{region "02 - Accept Start"}
// Accept Start into Starting; processing and Assertion evaluation are not active yet.
FSteps[2].RequestStart := TRUE;
FSteps[2].ExpectedState := E_State.Starting;
FSteps[2].ExpectedResult := E_Result.NotEvaluated;
FSteps[2].ExpectedReady := FALSE;
FSteps[2].ExpectedPassedCount := 0;
FSteps[2].ExpectedFailedCount := 0;
FSteps[2].ExpectedHookCount := 5;
FSteps[2].ExpectedHooks[1].Hook := E_LifecycleHook.Abort;
FSteps[2].ExpectedHooks[1].State := E_State.Starting;
FSteps[2].ExpectedHooks[1].Enabled := FALSE;
FSteps[2].ExpectedHooks[2].Hook := E_LifecycleHook.Preparations;
FSteps[2].ExpectedHooks[2].State := E_State.Starting;
FSteps[2].ExpectedHooks[2].Enabled := FALSE;
FSteps[2].ExpectedHooks[3].Hook := E_LifecycleHook.Tests;
FSteps[2].ExpectedHooks[3].State := E_State.Starting;
FSteps[2].ExpectedHooks[3].Enabled := FALSE;
FSteps[2].ExpectedHooks[4].Hook := E_LifecycleHook.Assertions;
FSteps[2].ExpectedHooks[4].State := E_State.Starting;
FSteps[2].ExpectedHooks[4].Enabled := FALSE;
FSteps[2].ExpectedHooks[5].Hook := E_LifecycleHook.Aggregate;
FSteps[2].ExpectedHooks[5].State := E_State.Starting;
FSteps[2].ExpectedHooks[5].Enabled := TRUE;
{endregion}

{region "03 - Enter Running"}
// Enter Running and evaluate both children; owner Result stays NotEvaluated until finalization.
FSteps[3].ExpectedState := E_State.Running;
FSteps[3].ExpectedResult := E_Result.NotEvaluated;
FSteps[3].ExpectedReady := FALSE;
FSteps[3].ExpectedPassedCount := 2;
FSteps[3].ExpectedFailedCount := 0;
FSteps[3].ExpectedHookCount := 5;
FSteps[3].ExpectedHooks[1].Hook := E_LifecycleHook.Abort;
FSteps[3].ExpectedHooks[1].State := E_State.Running;
FSteps[3].ExpectedHooks[1].Enabled := FALSE;
FSteps[3].ExpectedHooks[2].Hook := E_LifecycleHook.Preparations;
FSteps[3].ExpectedHooks[2].State := E_State.Running;
FSteps[3].ExpectedHooks[2].Enabled := FALSE;
FSteps[3].ExpectedHooks[3].Hook := E_LifecycleHook.Tests;
FSteps[3].ExpectedHooks[3].State := E_State.Running;
FSteps[3].ExpectedHooks[3].Enabled := TRUE;
FSteps[3].ExpectedHooks[4].Hook := E_LifecycleHook.Assertions;
FSteps[3].ExpectedHooks[4].State := E_State.Running;
FSteps[3].ExpectedHooks[4].Enabled := TRUE;
FSteps[3].ExpectedHooks[5].Hook := E_LifecycleHook.Aggregate;
FSteps[3].ExpectedHooks[5].State := E_State.Running;
FSteps[3].ExpectedHooks[5].Enabled := TRUE;
{endregion}

{region "04 - Request Abort and hold acknowledgement"}
// Request Abort once and withhold cleanup acknowledgement.
FSteps[4].RequestAbort := TRUE;
FSteps[4].AbortCompleted := FALSE;
FSteps[4].ExpectedState := E_State.Aborting;
FSteps[4].ExpectedResult := E_Result.Abort;
FSteps[4].ExpectedReady := FALSE;
FSteps[4].ExpectedPassedCount := 2;
FSteps[4].ExpectedFailedCount := 0;
FSteps[4].ExpectedHookCount := 5;
FSteps[4].ExpectedHooks[1].Hook := E_LifecycleHook.Abort;
FSteps[4].ExpectedHooks[1].State := E_State.Aborting;
FSteps[4].ExpectedHooks[1].Enabled := TRUE;
FSteps[4].ExpectedHooks[2].Hook := E_LifecycleHook.Preparations;
FSteps[4].ExpectedHooks[2].State := E_State.Aborting;
FSteps[4].ExpectedHooks[2].Enabled := FALSE;
FSteps[4].ExpectedHooks[3].Hook := E_LifecycleHook.Tests;
FSteps[4].ExpectedHooks[3].State := E_State.Aborting;
FSteps[4].ExpectedHooks[3].Enabled := FALSE;
FSteps[4].ExpectedHooks[4].Hook := E_LifecycleHook.Assertions;
FSteps[4].ExpectedHooks[4].State := E_State.Aborting;
FSteps[4].ExpectedHooks[4].Enabled := FALSE;
FSteps[4].ExpectedHooks[5].Hook := E_LifecycleHook.Aggregate;
FSteps[4].ExpectedHooks[5].State := E_State.Aborting;
FSteps[4].ExpectedHooks[5].Enabled := TRUE;
{endregion}

{region "05 - Wait for Abort timeout"}
// Keep cleanup open while repeating this checkpoint in Aborting.
// Timeout forces Completing with Error even though the implementation never acknowledges Abort.
FSteps[5].WaitForTransition := TRUE;
FSteps[5].WaitingState := E_State.Aborting;
FSteps[5].AbortCompleted := FALSE;
FSteps[5].ExpectedAbortTimeout := TRUE;
FSteps[5].ExpectedState := E_State.Completing;
FSteps[5].ExpectedResult := E_Result.Error;
FSteps[5].ExpectedReady := FALSE;
FSteps[5].ExpectedPassedCount := 2;
FSteps[5].ExpectedFailedCount := 0;
FSteps[5].ExpectedHookCount := 5;
FSteps[5].ExpectedHooks[1].Hook := E_LifecycleHook.Abort;
FSteps[5].ExpectedHooks[1].State := E_State.Completing;
FSteps[5].ExpectedHooks[1].Enabled := FALSE;
FSteps[5].ExpectedHooks[2].Hook := E_LifecycleHook.Preparations;
FSteps[5].ExpectedHooks[2].State := E_State.Completing;
FSteps[5].ExpectedHooks[2].Enabled := FALSE;
FSteps[5].ExpectedHooks[3].Hook := E_LifecycleHook.Tests;
FSteps[5].ExpectedHooks[3].State := E_State.Completing;
FSteps[5].ExpectedHooks[3].Enabled := FALSE;
FSteps[5].ExpectedHooks[4].Hook := E_LifecycleHook.Assertions;
FSteps[5].ExpectedHooks[4].State := E_State.Completing;
FSteps[5].ExpectedHooks[4].Enabled := FALSE;
FSteps[5].ExpectedHooks[5].Hook := E_LifecycleHook.Aggregate;
FSteps[5].ExpectedHooks[5].State := E_State.Completing;
FSteps[5].ExpectedHooks[5].Enabled := TRUE;
{endregion}

{region "06 - Retain timeout at completion"}
// Reach Completed and retain the Abort-timeout diagnostic.
FSteps[6].ExpectedAbortTimeout := TRUE;
FSteps[6].ExpectedState := E_State.Completed;
FSteps[6].ExpectedResult := E_Result.Error;
FSteps[6].ExpectedReady := FALSE;
FSteps[6].ExpectedPassedCount := 2;
FSteps[6].ExpectedFailedCount := 0;
FSteps[6].ExpectedHookCount := 1;
FSteps[6].ExpectedHooks[1].Hook := E_LifecycleHook.Aggregate;
FSteps[6].ExpectedHooks[1].State := E_State.Completed;
FSteps[6].ExpectedHooks[1].Enabled := TRUE;
{endregion}

{region "07 - Reset clears held timeout and result"}
FSteps[7].ExpectedState := E_State.Idle;
FSteps[7].ExpectedResult := E_Result.NotEvaluated;
FSteps[7].ExpectedReady := TRUE;
FSteps[7].ExpectedPassedCount := 0;
FSteps[7].ExpectedFailedCount := 0;
FSteps[7].CheckFinalization := TRUE;
FSteps[7].ExpectedFinalizationCount := 1;
FSteps[7].ExpectedCompletionCount := 1;
FSteps[7].ExpectedFinalResult := E_Result.Error;
FSteps[7].RequestReset := TRUE;
FSteps[7].PreparationTargetReached := TRUE;
FSteps[7].ExpectRuntimeCleared := TRUE;
FSteps[7].ExpectedHookCount := 6;
FSteps[7].ExpectedHooks[1].Hook := E_LifecycleHook.Reset;
FSteps[7].ExpectedHooks[1].State := E_State.Reset;
FSteps[7].ExpectedHooks[1].Enabled := TRUE;
FSteps[7].ExpectedHooks[2].Hook := E_LifecycleHook.Abort;
FSteps[7].ExpectedHooks[2].State := E_State.Idle;
FSteps[7].ExpectedHooks[2].Enabled := FALSE;
FSteps[7].ExpectedHooks[3].Hook := E_LifecycleHook.Preparations;
FSteps[7].ExpectedHooks[3].State := E_State.Idle;
FSteps[7].ExpectedHooks[3].Enabled := FALSE;
FSteps[7].ExpectedHooks[4].Hook := E_LifecycleHook.Tests;
FSteps[7].ExpectedHooks[4].State := E_State.Idle;
FSteps[7].ExpectedHooks[4].Enabled := FALSE;
FSteps[7].ExpectedHooks[5].Hook := E_LifecycleHook.Assertions;
FSteps[7].ExpectedHooks[5].State := E_State.Idle;
FSteps[7].ExpectedHooks[5].Enabled := FALSE;
FSteps[7].ExpectedHooks[6].Hook := E_LifecycleHook.Aggregate;
FSteps[7].ExpectedHooks[6].State := E_State.Idle;
FSteps[7].ExpectedHooks[6].Enabled := TRUE;
{endregion}

{region "08 - Start after timeout recovery"}
FSteps[8].ExpectedState := E_State.Starting;
FSteps[8].ExpectedResult := E_Result.NotEvaluated;
FSteps[8].ExpectedReady := FALSE;
FSteps[8].ExpectedPassedCount := 0;
FSteps[8].ExpectedFailedCount := 0;
FSteps[8].CheckFinalization := TRUE;
FSteps[8].ExpectedFinalizationCount := 1;
FSteps[8].ExpectedCompletionCount := 1;
FSteps[8].ExpectedFinalResult := E_Result.Error;
FSteps[8].RequestStart := TRUE;
FSteps[8].PreparationTargetReached := TRUE;
FSteps[8].ExpectedHookCount := 5;
FSteps[8].ExpectedHooks[1].Hook := E_LifecycleHook.Abort;
FSteps[8].ExpectedHooks[1].State := E_State.Starting;
FSteps[8].ExpectedHooks[1].Enabled := FALSE;
FSteps[8].ExpectedHooks[2].Hook := E_LifecycleHook.Preparations;
FSteps[8].ExpectedHooks[2].State := E_State.Starting;
FSteps[8].ExpectedHooks[2].Enabled := FALSE;
FSteps[8].ExpectedHooks[3].Hook := E_LifecycleHook.Tests;
FSteps[8].ExpectedHooks[3].State := E_State.Starting;
FSteps[8].ExpectedHooks[3].Enabled := FALSE;
FSteps[8].ExpectedHooks[4].Hook := E_LifecycleHook.Assertions;
FSteps[8].ExpectedHooks[4].State := E_State.Starting;
FSteps[8].ExpectedHooks[4].Enabled := FALSE;
FSteps[8].ExpectedHooks[5].Hook := E_LifecycleHook.Aggregate;
FSteps[8].ExpectedHooks[5].State := E_State.Starting;
FSteps[8].ExpectedHooks[5].Enabled := TRUE;
{endregion}

{region "09 - Execute without previous timeout flags"}
FSteps[9].ExpectedState := E_State.Running;
FSteps[9].ExpectedResult := E_Result.NotEvaluated;
FSteps[9].ExpectedReady := FALSE;
FSteps[9].ExpectedPassedCount := 2;
FSteps[9].ExpectedFailedCount := 0;
FSteps[9].CheckFinalization := TRUE;
FSteps[9].ExpectedFinalizationCount := 1;
FSteps[9].ExpectedCompletionCount := 1;
FSteps[9].ExpectedFinalResult := E_Result.Error;
FSteps[9].ExpectedHookCount := 5;
FSteps[9].ExpectedHooks[1].Hook := E_LifecycleHook.Abort;
FSteps[9].ExpectedHooks[1].State := E_State.Running;
FSteps[9].ExpectedHooks[1].Enabled := FALSE;
FSteps[9].ExpectedHooks[2].Hook := E_LifecycleHook.Preparations;
FSteps[9].ExpectedHooks[2].State := E_State.Running;
FSteps[9].ExpectedHooks[2].Enabled := FALSE;
FSteps[9].ExpectedHooks[3].Hook := E_LifecycleHook.Tests;
FSteps[9].ExpectedHooks[3].State := E_State.Running;
FSteps[9].ExpectedHooks[3].Enabled := TRUE;
FSteps[9].ExpectedHooks[4].Hook := E_LifecycleHook.Assertions;
FSteps[9].ExpectedHooks[4].State := E_State.Running;
FSteps[9].ExpectedHooks[4].Enabled := TRUE;
FSteps[9].ExpectedHooks[5].Hook := E_LifecycleHook.Aggregate;
FSteps[9].ExpectedHooks[5].State := E_State.Running;
FSteps[9].ExpectedHooks[5].Enabled := TRUE;
{endregion}

{region "10 - Finalize the recovered run"}
FSteps[10].ExpectedState := E_State.Completing;
FSteps[10].ExpectedResult := E_Result.Passed;
FSteps[10].ExpectedReady := FALSE;
FSteps[10].ExpectedPassedCount := 2;
FSteps[10].ExpectedFailedCount := 0;
FSteps[10].FinishTests := TRUE;
FSteps[10].CheckFinalization := TRUE;
FSteps[10].ExpectedFinalizationCount := 2;
FSteps[10].ExpectedCompletionCount := 1;
FSteps[10].ExpectedFinalResult := E_Result.Passed;
FSteps[10].ExpectedHookCount := 5;
FSteps[10].ExpectedHooks[1].Hook := E_LifecycleHook.Abort;
FSteps[10].ExpectedHooks[1].State := E_State.Running;
FSteps[10].ExpectedHooks[1].Enabled := FALSE;
FSteps[10].ExpectedHooks[2].Hook := E_LifecycleHook.Preparations;
FSteps[10].ExpectedHooks[2].State := E_State.Running;
FSteps[10].ExpectedHooks[2].Enabled := FALSE;
FSteps[10].ExpectedHooks[3].Hook := E_LifecycleHook.Tests;
FSteps[10].ExpectedHooks[3].State := E_State.Running;
FSteps[10].ExpectedHooks[3].Enabled := TRUE;
FSteps[10].ExpectedHooks[4].Hook := E_LifecycleHook.Assertions;
FSteps[10].ExpectedHooks[4].State := E_State.Completing;
FSteps[10].ExpectedHooks[4].Enabled := FALSE;
FSteps[10].ExpectedHooks[5].Hook := E_LifecycleHook.Aggregate;
FSteps[10].ExpectedHooks[5].State := E_State.Completing;
FSteps[10].ExpectedHooks[5].Enabled := TRUE;
{endregion}

{region "11 - Complete the recovered run"}
FSteps[11].ExpectedState := E_State.Completed;
FSteps[11].ExpectedResult := E_Result.Passed;
FSteps[11].ExpectedReady := FALSE;
FSteps[11].ExpectedPassedCount := 2;
FSteps[11].ExpectedFailedCount := 0;
FSteps[11].ExpectRuntimeHeld := TRUE;
FSteps[11].CheckFinalization := TRUE;
FSteps[11].ExpectedFinalizationCount := 2;
FSteps[11].ExpectedCompletionCount := 2;
FSteps[11].ExpectedFinalResult := E_Result.Passed;
FSteps[11].ExpectedHookCount := 1;
FSteps[11].ExpectedHooks[1].Hook := E_LifecycleHook.Aggregate;
FSteps[11].ExpectedHooks[1].State := E_State.Completed;
FSteps[11].ExpectedHooks[1].Enabled := TRUE;
{endregion}

{region "12 - Hold the recovered completion without new events"}
FSteps[12].ExpectedState := E_State.Completed;
FSteps[12].ExpectedResult := E_Result.Passed;
FSteps[12].ExpectedReady := FALSE;
FSteps[12].ExpectedPassedCount := 2;
FSteps[12].ExpectedFailedCount := 0;
FSteps[12].ExpectQuietCall := TRUE;
FSteps[12].ExpectRuntimeHeld := TRUE;
FSteps[12].CheckFinalization := TRUE;
FSteps[12].ExpectedFinalizationCount := 2;
FSteps[12].ExpectedCompletionCount := 2;
FSteps[12].ExpectedFinalResult := E_Result.Passed;
FSteps[12].ExpectedHookCount := 1;
FSteps[12].ExpectedHooks[1].Hook := E_LifecycleHook.Aggregate;
FSteps[12].ExpectedHooks[1].State := E_State.Completed;
FSteps[12].ExpectedHooks[1].Enabled := TRUE;
{endregion}
END_METHOD

END_FUNCTION_BLOCK

// ---- SelfTests/TestCases/TestSuite_TestCaseLifecycle/Test_LifecycleExecutionTimeout.TcPOU
{region 'Documentation'}
(*!
<summary>Leaves the Test phase pending until the real configured execution timeout finalizes Error.</summary>
*)
{endregion}
FUNCTION_BLOCK Test_LifecycleExecutionTimeout EXTENDS TestCaseLifecycleTestBase

SUPER^();

{region 'Documentation'}
(*!
<summary>Defines explicit exceptional-path stimuli and contract-derived observations.</summary>
*)
{endregion}
METHOD PROTECTED ConfigureScenario
// Exercise the real cyclic timer; these checkpoints check the timeout path and retained flag,
// not an exact elapsed-time boundary. The outer Test Case timeout bounds a missing transition.
FSubjectPreparationCount := 0;
FSubjectTestCount := 1;
FStepCount := 11;
FSubjectConfig.Timeout := T#50ms;

{region "01 - Reset to Idle"}
// Establish Idle through the parent Reset request; both child results must be cleared.
FSteps[1].RequestReset := TRUE;
FSteps[1].ExpectedState := E_State.Idle;
FSteps[1].ExpectedResult := E_Result.NotEvaluated;
FSteps[1].ExpectedReady := TRUE;
FSteps[1].ExpectedPassedCount := 0;
FSteps[1].ExpectedFailedCount := 0;
FSteps[1].ExpectedHookCount := 6;
FSteps[1].ExpectedHooks[1].Hook := E_LifecycleHook.Reset;
FSteps[1].ExpectedHooks[1].State := E_State.Reset;
FSteps[1].ExpectedHooks[1].Enabled := TRUE;
FSteps[1].ExpectedHooks[2].Hook := E_LifecycleHook.Abort;
FSteps[1].ExpectedHooks[2].State := E_State.Idle;
FSteps[1].ExpectedHooks[2].Enabled := FALSE;
FSteps[1].ExpectedHooks[3].Hook := E_LifecycleHook.Preparations;
FSteps[1].ExpectedHooks[3].State := E_State.Idle;
FSteps[1].ExpectedHooks[3].Enabled := FALSE;
FSteps[1].ExpectedHooks[4].Hook := E_LifecycleHook.Tests;
FSteps[1].ExpectedHooks[4].State := E_State.Idle;
FSteps[1].ExpectedHooks[4].Enabled := FALSE;
FSteps[1].ExpectedHooks[5].Hook := E_LifecycleHook.Assertions;
FSteps[1].ExpectedHooks[5].State := E_State.Idle;
FSteps[1].ExpectedHooks[5].Enabled := FALSE;
FSteps[1].ExpectedHooks[6].Hook := E_LifecycleHook.Aggregate;
FSteps[1].ExpectedHooks[6].State := E_State.Idle;
FSteps[1].ExpectedHooks[6].Enabled := TRUE;
{endregion}

{region "02 - Accept Start"}
// Accept Start into Starting; processing and Assertion evaluation are not active yet.
FSteps[2].RequestStart := TRUE;
FSteps[2].ExpectedState := E_State.Starting;
FSteps[2].ExpectedResult := E_Result.NotEvaluated;
FSteps[2].ExpectedReady := FALSE;
FSteps[2].ExpectedPassedCount := 0;
FSteps[2].ExpectedFailedCount := 0;
FSteps[2].ExpectedHookCount := 5;
FSteps[2].ExpectedHooks[1].Hook := E_LifecycleHook.Abort;
FSteps[2].ExpectedHooks[1].State := E_State.Starting;
FSteps[2].ExpectedHooks[1].Enabled := FALSE;
FSteps[2].ExpectedHooks[2].Hook := E_LifecycleHook.Preparations;
FSteps[2].ExpectedHooks[2].State := E_State.Starting;
FSteps[2].ExpectedHooks[2].Enabled := FALSE;
FSteps[2].ExpectedHooks[3].Hook := E_LifecycleHook.Tests;
FSteps[2].ExpectedHooks[3].State := E_State.Starting;
FSteps[2].ExpectedHooks[3].Enabled := FALSE;
FSteps[2].ExpectedHooks[4].Hook := E_LifecycleHook.Assertions;
FSteps[2].ExpectedHooks[4].State := E_State.Starting;
FSteps[2].ExpectedHooks[4].Enabled := FALSE;
FSteps[2].ExpectedHooks[5].Hook := E_LifecycleHook.Aggregate;
FSteps[2].ExpectedHooks[5].State := E_State.Starting;
FSteps[2].ExpectedHooks[5].Enabled := TRUE;
{endregion}

{region "03 - Enter Running"}
// Enter Running and evaluate both children; owner Result stays NotEvaluated until finalization.
FSteps[3].ExpectedState := E_State.Running;
FSteps[3].ExpectedResult := E_Result.NotEvaluated;
FSteps[3].ExpectedReady := FALSE;
FSteps[3].ExpectedPassedCount := 2;
FSteps[3].ExpectedFailedCount := 0;
FSteps[3].ExpectedHookCount := 5;
FSteps[3].ExpectedHooks[1].Hook := E_LifecycleHook.Abort;
FSteps[3].ExpectedHooks[1].State := E_State.Running;
FSteps[3].ExpectedHooks[1].Enabled := FALSE;
FSteps[3].ExpectedHooks[2].Hook := E_LifecycleHook.Preparations;
FSteps[3].ExpectedHooks[2].State := E_State.Running;
FSteps[3].ExpectedHooks[2].Enabled := FALSE;
FSteps[3].ExpectedHooks[3].Hook := E_LifecycleHook.Tests;
FSteps[3].ExpectedHooks[3].State := E_State.Running;
FSteps[3].ExpectedHooks[3].Enabled := TRUE;
FSteps[3].ExpectedHooks[4].Hook := E_LifecycleHook.Assertions;
FSteps[3].ExpectedHooks[4].State := E_State.Running;
FSteps[3].ExpectedHooks[4].Enabled := TRUE;
FSteps[3].ExpectedHooks[5].Hook := E_LifecycleHook.Aggregate;
FSteps[3].ExpectedHooks[5].State := E_State.Running;
FSteps[3].ExpectedHooks[5].Enabled := TRUE;
{endregion}

{region "04 - Wait for execution timeout"}
// Keep execution open and repeat this checkpoint while Running.
// On timeout, immediate abort cleanup reaches Completing with Error and HasTimeout set.
FSteps[4].WaitForTransition := TRUE;
FSteps[4].WaitingState := E_State.Running;
FSteps[4].ExpectedTimeout := TRUE;
FSteps[4].ExpectedState := E_State.Completing;
FSteps[4].ExpectedResult := E_Result.Error;
FSteps[4].ExpectedReady := FALSE;
FSteps[4].ExpectedPassedCount := 2;
FSteps[4].ExpectedFailedCount := 0;
FSteps[4].ExpectedHookCount := 5;
FSteps[4].ExpectedHooks[1].Hook := E_LifecycleHook.Abort;
FSteps[4].ExpectedHooks[1].State := E_State.AbortingFromError;
FSteps[4].ExpectedHooks[1].Enabled := TRUE;
FSteps[4].ExpectedHooks[2].Hook := E_LifecycleHook.Preparations;
FSteps[4].ExpectedHooks[2].State := E_State.Completing;
FSteps[4].ExpectedHooks[2].Enabled := FALSE;
FSteps[4].ExpectedHooks[3].Hook := E_LifecycleHook.Tests;
FSteps[4].ExpectedHooks[3].State := E_State.Completing;
FSteps[4].ExpectedHooks[3].Enabled := FALSE;
FSteps[4].ExpectedHooks[4].Hook := E_LifecycleHook.Assertions;
FSteps[4].ExpectedHooks[4].State := E_State.Completing;
FSteps[4].ExpectedHooks[4].Enabled := FALSE;
FSteps[4].ExpectedHooks[5].Hook := E_LifecycleHook.Aggregate;
FSteps[4].ExpectedHooks[5].State := E_State.Completing;
FSteps[4].ExpectedHooks[5].Enabled := TRUE;
{endregion}

{region "05 - Retain timeout at completion"}
// Reach Completed and retain the execution-timeout diagnostic.
FSteps[5].ExpectedTimeout := TRUE;
FSteps[5].ExpectedState := E_State.Completed;
FSteps[5].ExpectedResult := E_Result.Error;
FSteps[5].ExpectedReady := FALSE;
FSteps[5].ExpectedPassedCount := 2;
FSteps[5].ExpectedFailedCount := 0;
FSteps[5].ExpectedHookCount := 1;
FSteps[5].ExpectedHooks[1].Hook := E_LifecycleHook.Aggregate;
FSteps[5].ExpectedHooks[1].State := E_State.Completed;
FSteps[5].ExpectedHooks[1].Enabled := TRUE;
{endregion}

{region "06 - Reset clears held timeout and result"}
FSteps[6].ExpectedState := E_State.Idle;
FSteps[6].ExpectedResult := E_Result.NotEvaluated;
FSteps[6].ExpectedReady := TRUE;
FSteps[6].ExpectedPassedCount := 0;
FSteps[6].ExpectedFailedCount := 0;
FSteps[6].CheckFinalization := TRUE;
FSteps[6].ExpectedFinalizationCount := 1;
FSteps[6].ExpectedCompletionCount := 1;
FSteps[6].ExpectedFinalResult := E_Result.Error;
FSteps[6].RequestReset := TRUE;
FSteps[6].PreparationTargetReached := TRUE;
FSteps[6].ExpectRuntimeCleared := TRUE;
FSteps[6].ExpectedHookCount := 6;
FSteps[6].ExpectedHooks[1].Hook := E_LifecycleHook.Reset;
FSteps[6].ExpectedHooks[1].State := E_State.Reset;
FSteps[6].ExpectedHooks[1].Enabled := TRUE;
FSteps[6].ExpectedHooks[2].Hook := E_LifecycleHook.Abort;
FSteps[6].ExpectedHooks[2].State := E_State.Idle;
FSteps[6].ExpectedHooks[2].Enabled := FALSE;
FSteps[6].ExpectedHooks[3].Hook := E_LifecycleHook.Preparations;
FSteps[6].ExpectedHooks[3].State := E_State.Idle;
FSteps[6].ExpectedHooks[3].Enabled := FALSE;
FSteps[6].ExpectedHooks[4].Hook := E_LifecycleHook.Tests;
FSteps[6].ExpectedHooks[4].State := E_State.Idle;
FSteps[6].ExpectedHooks[4].Enabled := FALSE;
FSteps[6].ExpectedHooks[5].Hook := E_LifecycleHook.Assertions;
FSteps[6].ExpectedHooks[5].State := E_State.Idle;
FSteps[6].ExpectedHooks[5].Enabled := FALSE;
FSteps[6].ExpectedHooks[6].Hook := E_LifecycleHook.Aggregate;
FSteps[6].ExpectedHooks[6].State := E_State.Idle;
FSteps[6].ExpectedHooks[6].Enabled := TRUE;
{endregion}

{region "07 - Start after timeout recovery"}
FSteps[7].ExpectedState := E_State.Starting;
FSteps[7].ExpectedResult := E_Result.NotEvaluated;
FSteps[7].ExpectedReady := FALSE;
FSteps[7].ExpectedPassedCount := 0;
FSteps[7].ExpectedFailedCount := 0;
FSteps[7].CheckFinalization := TRUE;
FSteps[7].ExpectedFinalizationCount := 1;
FSteps[7].ExpectedCompletionCount := 1;
FSteps[7].ExpectedFinalResult := E_Result.Error;
FSteps[7].RequestStart := TRUE;
FSteps[7].PreparationTargetReached := TRUE;
FSteps[7].ExpectedHookCount := 5;
FSteps[7].ExpectedHooks[1].Hook := E_LifecycleHook.Abort;
FSteps[7].ExpectedHooks[1].State := E_State.Starting;
FSteps[7].ExpectedHooks[1].Enabled := FALSE;
FSteps[7].ExpectedHooks[2].Hook := E_LifecycleHook.Preparations;
FSteps[7].ExpectedHooks[2].State := E_State.Starting;
FSteps[7].ExpectedHooks[2].Enabled := FALSE;
FSteps[7].ExpectedHooks[3].Hook := E_LifecycleHook.Tests;
FSteps[7].ExpectedHooks[3].State := E_State.Starting;
FSteps[7].ExpectedHooks[3].Enabled := FALSE;
FSteps[7].ExpectedHooks[4].Hook := E_LifecycleHook.Assertions;
FSteps[7].ExpectedHooks[4].State := E_State.Starting;
FSteps[7].ExpectedHooks[4].Enabled := FALSE;
FSteps[7].ExpectedHooks[5].Hook := E_LifecycleHook.Aggregate;
FSteps[7].ExpectedHooks[5].State := E_State.Starting;
FSteps[7].ExpectedHooks[5].Enabled := TRUE;
{endregion}

{region "08 - Execute without previous timeout flags"}
FSteps[8].ExpectedState := E_State.Running;
FSteps[8].ExpectedResult := E_Result.NotEvaluated;
FSteps[8].ExpectedReady := FALSE;
FSteps[8].ExpectedPassedCount := 2;
FSteps[8].ExpectedFailedCount := 0;
FSteps[8].CheckFinalization := TRUE;
FSteps[8].ExpectedFinalizationCount := 1;
FSteps[8].ExpectedCompletionCount := 1;
FSteps[8].ExpectedFinalResult := E_Result.Error;
FSteps[8].ExpectedHookCount := 5;
FSteps[8].ExpectedHooks[1].Hook := E_LifecycleHook.Abort;
FSteps[8].ExpectedHooks[1].State := E_State.Running;
FSteps[8].ExpectedHooks[1].Enabled := FALSE;
FSteps[8].ExpectedHooks[2].Hook := E_LifecycleHook.Preparations;
FSteps[8].ExpectedHooks[2].State := E_State.Running;
FSteps[8].ExpectedHooks[2].Enabled := FALSE;
FSteps[8].ExpectedHooks[3].Hook := E_LifecycleHook.Tests;
FSteps[8].ExpectedHooks[3].State := E_State.Running;
FSteps[8].ExpectedHooks[3].Enabled := TRUE;
FSteps[8].ExpectedHooks[4].Hook := E_LifecycleHook.Assertions;
FSteps[8].ExpectedHooks[4].State := E_State.Running;
FSteps[8].ExpectedHooks[4].Enabled := TRUE;
FSteps[8].ExpectedHooks[5].Hook := E_LifecycleHook.Aggregate;
FSteps[8].ExpectedHooks[5].State := E_State.Running;
FSteps[8].ExpectedHooks[5].Enabled := TRUE;
{endregion}

{region "09 - Finalize the recovered run"}
FSteps[9].ExpectedState := E_State.Completing;
FSteps[9].ExpectedResult := E_Result.Passed;
FSteps[9].ExpectedReady := FALSE;
FSteps[9].ExpectedPassedCount := 2;
FSteps[9].ExpectedFailedCount := 0;
FSteps[9].FinishTests := TRUE;
FSteps[9].CheckFinalization := TRUE;
FSteps[9].ExpectedFinalizationCount := 2;
FSteps[9].ExpectedCompletionCount := 1;
FSteps[9].ExpectedFinalResult := E_Result.Passed;
FSteps[9].ExpectedHookCount := 5;
FSteps[9].ExpectedHooks[1].Hook := E_LifecycleHook.Abort;
FSteps[9].ExpectedHooks[1].State := E_State.Running;
FSteps[9].ExpectedHooks[1].Enabled := FALSE;
FSteps[9].ExpectedHooks[2].Hook := E_LifecycleHook.Preparations;
FSteps[9].ExpectedHooks[2].State := E_State.Running;
FSteps[9].ExpectedHooks[2].Enabled := FALSE;
FSteps[9].ExpectedHooks[3].Hook := E_LifecycleHook.Tests;
FSteps[9].ExpectedHooks[3].State := E_State.Running;
FSteps[9].ExpectedHooks[3].Enabled := TRUE;
FSteps[9].ExpectedHooks[4].Hook := E_LifecycleHook.Assertions;
FSteps[9].ExpectedHooks[4].State := E_State.Completing;
FSteps[9].ExpectedHooks[4].Enabled := FALSE;
FSteps[9].ExpectedHooks[5].Hook := E_LifecycleHook.Aggregate;
FSteps[9].ExpectedHooks[5].State := E_State.Completing;
FSteps[9].ExpectedHooks[5].Enabled := TRUE;
{endregion}

{region "10 - Complete the recovered run"}
FSteps[10].ExpectedState := E_State.Completed;
FSteps[10].ExpectedResult := E_Result.Passed;
FSteps[10].ExpectedReady := FALSE;
FSteps[10].ExpectedPassedCount := 2;
FSteps[10].ExpectedFailedCount := 0;
FSteps[10].ExpectRuntimeHeld := TRUE;
FSteps[10].CheckFinalization := TRUE;
FSteps[10].ExpectedFinalizationCount := 2;
FSteps[10].ExpectedCompletionCount := 2;
FSteps[10].ExpectedFinalResult := E_Result.Passed;
FSteps[10].ExpectedHookCount := 1;
FSteps[10].ExpectedHooks[1].Hook := E_LifecycleHook.Aggregate;
FSteps[10].ExpectedHooks[1].State := E_State.Completed;
FSteps[10].ExpectedHooks[1].Enabled := TRUE;
{endregion}

{region "11 - Hold the recovered completion without new events"}
FSteps[11].ExpectedState := E_State.Completed;
FSteps[11].ExpectedResult := E_Result.Passed;
FSteps[11].ExpectedReady := FALSE;
FSteps[11].ExpectedPassedCount := 2;
FSteps[11].ExpectedFailedCount := 0;
FSteps[11].ExpectQuietCall := TRUE;
FSteps[11].ExpectRuntimeHeld := TRUE;
FSteps[11].CheckFinalization := TRUE;
FSteps[11].ExpectedFinalizationCount := 2;
FSteps[11].ExpectedCompletionCount := 2;
FSteps[11].ExpectedFinalResult := E_Result.Passed;
FSteps[11].ExpectedHookCount := 1;
FSteps[11].ExpectedHooks[1].Hook := E_LifecycleHook.Aggregate;
FSteps[11].ExpectedHooks[1].State := E_State.Completed;
FSteps[11].ExpectedHooks[1].Enabled := TRUE;
{endregion}
END_METHOD

END_FUNCTION_BLOCK

// ---- SelfTests/TestCases/TestSuite_TestCaseLifecycle/Test_LifecyclePreparationError.TcPOU
{region 'Documentation'}
(*!
<summary>Checks that an observed Preparation error prevents all enabled Test calls.</summary>
*)
{endregion}
FUNCTION_BLOCK Test_LifecyclePreparationError EXTENDS TestCaseLifecycleTestBase

SUPER^();

{region 'Documentation'}
(*!
<summary>Defines explicit exceptional-path stimuli and contract-derived observations.</summary>
*)
{endregion}
METHOD PROTECTED ConfigureScenario
FSubjectPreparationCount := 1;
FSubjectTestCount := 1;
FStepCount := 5;

{region "01 - Reset to Idle"}
// Establish Idle through the parent Reset request; both child results must be cleared.
FSteps[1].RequestReset := TRUE;
FSteps[1].ExpectedState := E_State.Idle;
FSteps[1].ExpectedResult := E_Result.NotEvaluated;
FSteps[1].ExpectedReady := TRUE;
FSteps[1].ExpectedPassedCount := 0;
FSteps[1].ExpectedFailedCount := 0;
FSteps[1].ExpectedHookCount := 6;
FSteps[1].ExpectedHooks[1].Hook := E_LifecycleHook.Reset;
FSteps[1].ExpectedHooks[1].State := E_State.Reset;
FSteps[1].ExpectedHooks[1].Enabled := TRUE;
FSteps[1].ExpectedHooks[2].Hook := E_LifecycleHook.Abort;
FSteps[1].ExpectedHooks[2].State := E_State.Idle;
FSteps[1].ExpectedHooks[2].Enabled := FALSE;
FSteps[1].ExpectedHooks[3].Hook := E_LifecycleHook.Preparations;
FSteps[1].ExpectedHooks[3].State := E_State.Idle;
FSteps[1].ExpectedHooks[3].Enabled := FALSE;
FSteps[1].ExpectedHooks[4].Hook := E_LifecycleHook.Tests;
FSteps[1].ExpectedHooks[4].State := E_State.Idle;
FSteps[1].ExpectedHooks[4].Enabled := FALSE;
FSteps[1].ExpectedHooks[5].Hook := E_LifecycleHook.Assertions;
FSteps[1].ExpectedHooks[5].State := E_State.Idle;
FSteps[1].ExpectedHooks[5].Enabled := FALSE;
FSteps[1].ExpectedHooks[6].Hook := E_LifecycleHook.Aggregate;
FSteps[1].ExpectedHooks[6].State := E_State.Idle;
FSteps[1].ExpectedHooks[6].Enabled := TRUE;
{endregion}

{region "02 - Accept Start"}
// Accept Start into Starting; processing and Assertion evaluation are not active yet.
FSteps[2].RequestStart := TRUE;
FSteps[2].ExpectedState := E_State.Starting;
FSteps[2].ExpectedResult := E_Result.NotEvaluated;
FSteps[2].ExpectedReady := FALSE;
FSteps[2].ExpectedPassedCount := 0;
FSteps[2].ExpectedFailedCount := 0;
FSteps[2].ExpectedHookCount := 5;
FSteps[2].ExpectedHooks[1].Hook := E_LifecycleHook.Abort;
FSteps[2].ExpectedHooks[1].State := E_State.Starting;
FSteps[2].ExpectedHooks[1].Enabled := FALSE;
FSteps[2].ExpectedHooks[2].Hook := E_LifecycleHook.Preparations;
FSteps[2].ExpectedHooks[2].State := E_State.Starting;
FSteps[2].ExpectedHooks[2].Enabled := FALSE;
FSteps[2].ExpectedHooks[3].Hook := E_LifecycleHook.Tests;
FSteps[2].ExpectedHooks[3].State := E_State.Starting;
FSteps[2].ExpectedHooks[3].Enabled := FALSE;
FSteps[2].ExpectedHooks[4].Hook := E_LifecycleHook.Assertions;
FSteps[2].ExpectedHooks[4].State := E_State.Starting;
FSteps[2].ExpectedHooks[4].Enabled := FALSE;
FSteps[2].ExpectedHooks[5].Hook := E_LifecycleHook.Aggregate;
FSteps[2].ExpectedHooks[5].State := E_State.Starting;
FSteps[2].ExpectedHooks[5].Enabled := TRUE;
{endregion}

{region "03 - Publish Preparation error"}
// Publish a Preparation error after the Sequencer ran; the current owner state remains
// Preparing.
FSteps[3].PreparationError := TRUE;
FSteps[3].ExpectedState := E_State.Preparing;
FSteps[3].ExpectedResult := E_Result.NotEvaluated;
FSteps[3].ExpectedReady := FALSE;
FSteps[3].ExpectedPassedCount := 0;
FSteps[3].ExpectedFailedCount := 0;
FSteps[3].ExpectedHookCount := 5;
FSteps[3].ExpectedHooks[1].Hook := E_LifecycleHook.Abort;
FSteps[3].ExpectedHooks[1].State := E_State.Preparing;
FSteps[3].ExpectedHooks[1].Enabled := FALSE;
FSteps[3].ExpectedHooks[2].Hook := E_LifecycleHook.Preparations;
FSteps[3].ExpectedHooks[2].State := E_State.Preparing;
FSteps[3].ExpectedHooks[2].Enabled := TRUE;
FSteps[3].ExpectedHooks[3].Hook := E_LifecycleHook.Tests;
FSteps[3].ExpectedHooks[3].State := E_State.Preparing;
FSteps[3].ExpectedHooks[3].Enabled := FALSE;
FSteps[3].ExpectedHooks[4].Hook := E_LifecycleHook.Assertions;
FSteps[3].ExpectedHooks[4].State := E_State.Preparing;
FSteps[3].ExpectedHooks[4].Enabled := FALSE;
FSteps[3].ExpectedHooks[5].Hook := E_LifecycleHook.Aggregate;
FSteps[3].ExpectedHooks[5].State := E_State.Preparing;
FSteps[3].ExpectedHooks[5].Enabled := TRUE;
{endregion}

{region "04 - Consume error before processing"}
// The next Sequencer consumes that error before processing hooks.
// Abort cleanup completes immediately, and test Assertions must never become enabled.
FSteps[4].ExpectedState := E_State.Completing;
FSteps[4].ExpectedResult := E_Result.Error;
FSteps[4].ExpectedReady := FALSE;
FSteps[4].ExpectedPassedCount := 0;
FSteps[4].ExpectedFailedCount := 0;
FSteps[4].ExpectedHookCount := 5;
FSteps[4].ExpectedHooks[1].Hook := E_LifecycleHook.Abort;
FSteps[4].ExpectedHooks[1].State := E_State.AbortingFromError;
FSteps[4].ExpectedHooks[1].Enabled := TRUE;
FSteps[4].ExpectedHooks[2].Hook := E_LifecycleHook.Preparations;
FSteps[4].ExpectedHooks[2].State := E_State.Completing;
FSteps[4].ExpectedHooks[2].Enabled := FALSE;
FSteps[4].ExpectedHooks[3].Hook := E_LifecycleHook.Tests;
FSteps[4].ExpectedHooks[3].State := E_State.Completing;
FSteps[4].ExpectedHooks[3].Enabled := FALSE;
FSteps[4].ExpectedHooks[4].Hook := E_LifecycleHook.Assertions;
FSteps[4].ExpectedHooks[4].State := E_State.Completing;
FSteps[4].ExpectedHooks[4].Enabled := FALSE;
FSteps[4].ExpectedHooks[5].Hook := E_LifecycleHook.Aggregate;
FSteps[4].ExpectedHooks[5].State := E_State.Completing;
FSteps[4].ExpectedHooks[5].Enabled := TRUE;
{endregion}

{region "05 - Observe terminal Error"}
// The following call reaches Completed; only aggregation remains in the recorded processing
// hooks.
FSteps[5].ExpectedState := E_State.Completed;
FSteps[5].ExpectedResult := E_Result.Error;
FSteps[5].ExpectedReady := FALSE;
FSteps[5].ExpectedPassedCount := 0;
FSteps[5].ExpectedFailedCount := 0;
FSteps[5].ExpectedHookCount := 1;
FSteps[5].ExpectedHooks[1].Hook := E_LifecycleHook.Aggregate;
FSteps[5].ExpectedHooks[1].State := E_State.Completed;
FSteps[5].ExpectedHooks[1].Enabled := TRUE;
{endregion}
END_METHOD

END_FUNCTION_BLOCK

// ---- SelfTests/TestCases/TestSuite_TestCaseLifecycle/Test_LifecyclePreparationTimeout.TcPOU
{region 'Documentation'}
(*!
<summary>Leaves Preparation incomplete until its real deadline, without entering the Test phase.</summary>
*)
{endregion}
FUNCTION_BLOCK Test_LifecyclePreparationTimeout EXTENDS TestCaseLifecycleTestBase

SUPER^();

{region 'Documentation'}
(*!
<summary>Defines explicit exceptional-path stimuli and contract-derived observations.</summary>
*)
{endregion}
METHOD PROTECTED ConfigureScenario
// Exercise the real cyclic timer; these checkpoints check the timeout path and retained flag,
// not an exact elapsed-time boundary. The outer Test Case timeout bounds a missing transition.
FSubjectPreparationCount := 1;
FSubjectTestCount := 1;
FStepCount := 11;
FSubjectConfig.PreparationTimeout := T#50ms;

{region "01 - Reset to Idle"}
// Establish Idle through the parent Reset request; both child results must be cleared.
FSteps[1].RequestReset := TRUE;
FSteps[1].ExpectedState := E_State.Idle;
FSteps[1].ExpectedResult := E_Result.NotEvaluated;
FSteps[1].ExpectedReady := TRUE;
FSteps[1].ExpectedPassedCount := 0;
FSteps[1].ExpectedFailedCount := 0;
FSteps[1].ExpectedHookCount := 6;
FSteps[1].ExpectedHooks[1].Hook := E_LifecycleHook.Reset;
FSteps[1].ExpectedHooks[1].State := E_State.Reset;
FSteps[1].ExpectedHooks[1].Enabled := TRUE;
FSteps[1].ExpectedHooks[2].Hook := E_LifecycleHook.Abort;
FSteps[1].ExpectedHooks[2].State := E_State.Idle;
FSteps[1].ExpectedHooks[2].Enabled := FALSE;
FSteps[1].ExpectedHooks[3].Hook := E_LifecycleHook.Preparations;
FSteps[1].ExpectedHooks[3].State := E_State.Idle;
FSteps[1].ExpectedHooks[3].Enabled := FALSE;
FSteps[1].ExpectedHooks[4].Hook := E_LifecycleHook.Tests;
FSteps[1].ExpectedHooks[4].State := E_State.Idle;
FSteps[1].ExpectedHooks[4].Enabled := FALSE;
FSteps[1].ExpectedHooks[5].Hook := E_LifecycleHook.Assertions;
FSteps[1].ExpectedHooks[5].State := E_State.Idle;
FSteps[1].ExpectedHooks[5].Enabled := FALSE;
FSteps[1].ExpectedHooks[6].Hook := E_LifecycleHook.Aggregate;
FSteps[1].ExpectedHooks[6].State := E_State.Idle;
FSteps[1].ExpectedHooks[6].Enabled := TRUE;
{endregion}

{region "02 - Accept Start"}
// Accept Start into Starting; processing and Assertion evaluation are not active yet.
FSteps[2].RequestStart := TRUE;
FSteps[2].ExpectedState := E_State.Starting;
FSteps[2].ExpectedResult := E_Result.NotEvaluated;
FSteps[2].ExpectedReady := FALSE;
FSteps[2].ExpectedPassedCount := 0;
FSteps[2].ExpectedFailedCount := 0;
FSteps[2].ExpectedHookCount := 5;
FSteps[2].ExpectedHooks[1].Hook := E_LifecycleHook.Abort;
FSteps[2].ExpectedHooks[1].State := E_State.Starting;
FSteps[2].ExpectedHooks[1].Enabled := FALSE;
FSteps[2].ExpectedHooks[2].Hook := E_LifecycleHook.Preparations;
FSteps[2].ExpectedHooks[2].State := E_State.Starting;
FSteps[2].ExpectedHooks[2].Enabled := FALSE;
FSteps[2].ExpectedHooks[3].Hook := E_LifecycleHook.Tests;
FSteps[2].ExpectedHooks[3].State := E_State.Starting;
FSteps[2].ExpectedHooks[3].Enabled := FALSE;
FSteps[2].ExpectedHooks[4].Hook := E_LifecycleHook.Assertions;
FSteps[2].ExpectedHooks[4].State := E_State.Starting;
FSteps[2].ExpectedHooks[4].Enabled := FALSE;
FSteps[2].ExpectedHooks[5].Hook := E_LifecycleHook.Aggregate;
FSteps[2].ExpectedHooks[5].State := E_State.Starting;
FSteps[2].ExpectedHooks[5].Enabled := TRUE;
{endregion}

{region "03 - Enter Preparing"}
// Enter Preparing without evaluating Assertions; the target has not been reached.
FSteps[3].ExpectedState := E_State.Preparing;
FSteps[3].ExpectedResult := E_Result.NotEvaluated;
FSteps[3].ExpectedReady := FALSE;
FSteps[3].ExpectedPassedCount := 0;
FSteps[3].ExpectedFailedCount := 0;
FSteps[3].ExpectedHookCount := 5;
FSteps[3].ExpectedHooks[1].Hook := E_LifecycleHook.Abort;
FSteps[3].ExpectedHooks[1].State := E_State.Preparing;
FSteps[3].ExpectedHooks[1].Enabled := FALSE;
FSteps[3].ExpectedHooks[2].Hook := E_LifecycleHook.Preparations;
FSteps[3].ExpectedHooks[2].State := E_State.Preparing;
FSteps[3].ExpectedHooks[2].Enabled := TRUE;
FSteps[3].ExpectedHooks[3].Hook := E_LifecycleHook.Tests;
FSteps[3].ExpectedHooks[3].State := E_State.Preparing;
FSteps[3].ExpectedHooks[3].Enabled := FALSE;
FSteps[3].ExpectedHooks[4].Hook := E_LifecycleHook.Assertions;
FSteps[3].ExpectedHooks[4].State := E_State.Preparing;
FSteps[3].ExpectedHooks[4].Enabled := FALSE;
FSteps[3].ExpectedHooks[5].Hook := E_LifecycleHook.Aggregate;
FSteps[3].ExpectedHooks[5].State := E_State.Preparing;
FSteps[3].ExpectedHooks[5].Enabled := TRUE;
{endregion}

{region "04 - Wait for Preparation timeout"}
// Never report the target reached; repeat while Preparing.
// Preparation timeout must finalize through abort cleanup without evaluating any Assertion.
FSteps[4].WaitForTransition := TRUE;
FSteps[4].WaitingState := E_State.Preparing;
FSteps[4].ExpectedPreparationTimeout := TRUE;
FSteps[4].ExpectedState := E_State.Completing;
FSteps[4].ExpectedResult := E_Result.Error;
FSteps[4].ExpectedReady := FALSE;
FSteps[4].ExpectedPassedCount := 0;
FSteps[4].ExpectedFailedCount := 0;
FSteps[4].ExpectedHookCount := 5;
FSteps[4].ExpectedHooks[1].Hook := E_LifecycleHook.Abort;
FSteps[4].ExpectedHooks[1].State := E_State.AbortingFromError;
FSteps[4].ExpectedHooks[1].Enabled := TRUE;
FSteps[4].ExpectedHooks[2].Hook := E_LifecycleHook.Preparations;
FSteps[4].ExpectedHooks[2].State := E_State.Completing;
FSteps[4].ExpectedHooks[2].Enabled := FALSE;
FSteps[4].ExpectedHooks[3].Hook := E_LifecycleHook.Tests;
FSteps[4].ExpectedHooks[3].State := E_State.Completing;
FSteps[4].ExpectedHooks[3].Enabled := FALSE;
FSteps[4].ExpectedHooks[4].Hook := E_LifecycleHook.Assertions;
FSteps[4].ExpectedHooks[4].State := E_State.Completing;
FSteps[4].ExpectedHooks[4].Enabled := FALSE;
FSteps[4].ExpectedHooks[5].Hook := E_LifecycleHook.Aggregate;
FSteps[4].ExpectedHooks[5].State := E_State.Completing;
FSteps[4].ExpectedHooks[5].Enabled := TRUE;
{endregion}

{region "05 - Retain timeout at completion"}
// Reach Completed and retain the Preparation-timeout diagnostic.
FSteps[5].ExpectedPreparationTimeout := TRUE;
FSteps[5].ExpectedState := E_State.Completed;
FSteps[5].ExpectedResult := E_Result.Error;
FSteps[5].ExpectedReady := FALSE;
FSteps[5].ExpectedPassedCount := 0;
FSteps[5].ExpectedFailedCount := 0;
FSteps[5].ExpectedHookCount := 1;
FSteps[5].ExpectedHooks[1].Hook := E_LifecycleHook.Aggregate;
FSteps[5].ExpectedHooks[1].State := E_State.Completed;
FSteps[5].ExpectedHooks[1].Enabled := TRUE;
{endregion}

{region "06 - Reset clears held timeout and result"}
FSteps[6].ExpectedState := E_State.Idle;
FSteps[6].ExpectedResult := E_Result.NotEvaluated;
FSteps[6].ExpectedReady := TRUE;
FSteps[6].ExpectedPassedCount := 0;
FSteps[6].ExpectedFailedCount := 0;
FSteps[6].CheckFinalization := TRUE;
FSteps[6].ExpectedFinalizationCount := 1;
FSteps[6].ExpectedCompletionCount := 1;
FSteps[6].ExpectedFinalResult := E_Result.Error;
FSteps[6].RequestReset := TRUE;
FSteps[6].PreparationTargetReached := TRUE;
FSteps[6].ExpectRuntimeCleared := TRUE;
FSteps[6].ExpectedHookCount := 6;
FSteps[6].ExpectedHooks[1].Hook := E_LifecycleHook.Reset;
FSteps[6].ExpectedHooks[1].State := E_State.Reset;
FSteps[6].ExpectedHooks[1].Enabled := TRUE;
FSteps[6].ExpectedHooks[2].Hook := E_LifecycleHook.Abort;
FSteps[6].ExpectedHooks[2].State := E_State.Idle;
FSteps[6].ExpectedHooks[2].Enabled := FALSE;
FSteps[6].ExpectedHooks[3].Hook := E_LifecycleHook.Preparations;
FSteps[6].ExpectedHooks[3].State := E_State.Idle;
FSteps[6].ExpectedHooks[3].Enabled := FALSE;
FSteps[6].ExpectedHooks[4].Hook := E_LifecycleHook.Tests;
FSteps[6].ExpectedHooks[4].State := E_State.Idle;
FSteps[6].ExpectedHooks[4].Enabled := FALSE;
FSteps[6].ExpectedHooks[5].Hook := E_LifecycleHook.Assertions;
FSteps[6].ExpectedHooks[5].State := E_State.Idle;
FSteps[6].ExpectedHooks[5].Enabled := FALSE;
FSteps[6].ExpectedHooks[6].Hook := E_LifecycleHook.Aggregate;
FSteps[6].ExpectedHooks[6].State := E_State.Idle;
FSteps[6].ExpectedHooks[6].Enabled := TRUE;
{endregion}

{region "07 - Start after timeout recovery"}
FSteps[7].ExpectedState := E_State.Starting;
FSteps[7].ExpectedResult := E_Result.NotEvaluated;
FSteps[7].ExpectedReady := FALSE;
FSteps[7].ExpectedPassedCount := 0;
FSteps[7].ExpectedFailedCount := 0;
FSteps[7].CheckFinalization := TRUE;
FSteps[7].ExpectedFinalizationCount := 1;
FSteps[7].ExpectedCompletionCount := 1;
FSteps[7].ExpectedFinalResult := E_Result.Error;
FSteps[7].RequestStart := TRUE;
FSteps[7].PreparationTargetReached := TRUE;
FSteps[7].ExpectedHookCount := 5;
FSteps[7].ExpectedHooks[1].Hook := E_LifecycleHook.Abort;
FSteps[7].ExpectedHooks[1].State := E_State.Starting;
FSteps[7].ExpectedHooks[1].Enabled := FALSE;
FSteps[7].ExpectedHooks[2].Hook := E_LifecycleHook.Preparations;
FSteps[7].ExpectedHooks[2].State := E_State.Starting;
FSteps[7].ExpectedHooks[2].Enabled := FALSE;
FSteps[7].ExpectedHooks[3].Hook := E_LifecycleHook.Tests;
FSteps[7].ExpectedHooks[3].State := E_State.Starting;
FSteps[7].ExpectedHooks[3].Enabled := FALSE;
FSteps[7].ExpectedHooks[4].Hook := E_LifecycleHook.Assertions;
FSteps[7].ExpectedHooks[4].State := E_State.Starting;
FSteps[7].ExpectedHooks[4].Enabled := FALSE;
FSteps[7].ExpectedHooks[5].Hook := E_LifecycleHook.Aggregate;
FSteps[7].ExpectedHooks[5].State := E_State.Starting;
FSteps[7].ExpectedHooks[5].Enabled := TRUE;
{endregion}

{region "08 - Execute without previous timeout flags"}
FSteps[8].ExpectedState := E_State.Running;
FSteps[8].ExpectedResult := E_Result.NotEvaluated;
FSteps[8].ExpectedReady := FALSE;
FSteps[8].ExpectedPassedCount := 2;
FSteps[8].ExpectedFailedCount := 0;
FSteps[8].CheckFinalization := TRUE;
FSteps[8].ExpectedFinalizationCount := 1;
FSteps[8].ExpectedCompletionCount := 1;
FSteps[8].ExpectedFinalResult := E_Result.Error;
FSteps[8].ExpectedHookCount := 5;
FSteps[8].ExpectedHooks[1].Hook := E_LifecycleHook.Abort;
FSteps[8].ExpectedHooks[1].State := E_State.Running;
FSteps[8].ExpectedHooks[1].Enabled := FALSE;
FSteps[8].ExpectedHooks[2].Hook := E_LifecycleHook.Preparations;
FSteps[8].ExpectedHooks[2].State := E_State.Running;
FSteps[8].ExpectedHooks[2].Enabled := FALSE;
FSteps[8].ExpectedHooks[3].Hook := E_LifecycleHook.Tests;
FSteps[8].ExpectedHooks[3].State := E_State.Running;
FSteps[8].ExpectedHooks[3].Enabled := TRUE;
FSteps[8].ExpectedHooks[4].Hook := E_LifecycleHook.Assertions;
FSteps[8].ExpectedHooks[4].State := E_State.Running;
FSteps[8].ExpectedHooks[4].Enabled := TRUE;
FSteps[8].ExpectedHooks[5].Hook := E_LifecycleHook.Aggregate;
FSteps[8].ExpectedHooks[5].State := E_State.Running;
FSteps[8].ExpectedHooks[5].Enabled := TRUE;
{endregion}

{region "09 - Finalize the recovered run"}
FSteps[9].ExpectedState := E_State.Completing;
FSteps[9].ExpectedResult := E_Result.Passed;
FSteps[9].ExpectedReady := FALSE;
FSteps[9].ExpectedPassedCount := 2;
FSteps[9].ExpectedFailedCount := 0;
FSteps[9].FinishTests := TRUE;
FSteps[9].CheckFinalization := TRUE;
FSteps[9].ExpectedFinalizationCount := 2;
FSteps[9].ExpectedCompletionCount := 1;
FSteps[9].ExpectedFinalResult := E_Result.Passed;
FSteps[9].ExpectedHookCount := 5;
FSteps[9].ExpectedHooks[1].Hook := E_LifecycleHook.Abort;
FSteps[9].ExpectedHooks[1].State := E_State.Running;
FSteps[9].ExpectedHooks[1].Enabled := FALSE;
FSteps[9].ExpectedHooks[2].Hook := E_LifecycleHook.Preparations;
FSteps[9].ExpectedHooks[2].State := E_State.Running;
FSteps[9].ExpectedHooks[2].Enabled := FALSE;
FSteps[9].ExpectedHooks[3].Hook := E_LifecycleHook.Tests;
FSteps[9].ExpectedHooks[3].State := E_State.Running;
FSteps[9].ExpectedHooks[3].Enabled := TRUE;
FSteps[9].ExpectedHooks[4].Hook := E_LifecycleHook.Assertions;
FSteps[9].ExpectedHooks[4].State := E_State.Completing;
FSteps[9].ExpectedHooks[4].Enabled := FALSE;
FSteps[9].ExpectedHooks[5].Hook := E_LifecycleHook.Aggregate;
FSteps[9].ExpectedHooks[5].State := E_State.Completing;
FSteps[9].ExpectedHooks[5].Enabled := TRUE;
{endregion}

{region "10 - Complete the recovered run"}
FSteps[10].ExpectedState := E_State.Completed;
FSteps[10].ExpectedResult := E_Result.Passed;
FSteps[10].ExpectedReady := FALSE;
FSteps[10].ExpectedPassedCount := 2;
FSteps[10].ExpectedFailedCount := 0;
FSteps[10].ExpectRuntimeHeld := TRUE;
FSteps[10].CheckFinalization := TRUE;
FSteps[10].ExpectedFinalizationCount := 2;
FSteps[10].ExpectedCompletionCount := 2;
FSteps[10].ExpectedFinalResult := E_Result.Passed;
FSteps[10].ExpectedHookCount := 1;
FSteps[10].ExpectedHooks[1].Hook := E_LifecycleHook.Aggregate;
FSteps[10].ExpectedHooks[1].State := E_State.Completed;
FSteps[10].ExpectedHooks[1].Enabled := TRUE;
{endregion}

{region "11 - Hold the recovered completion without new events"}
FSteps[11].ExpectedState := E_State.Completed;
FSteps[11].ExpectedResult := E_Result.Passed;
FSteps[11].ExpectedReady := FALSE;
FSteps[11].ExpectedPassedCount := 2;
FSteps[11].ExpectedFailedCount := 0;
FSteps[11].ExpectQuietCall := TRUE;
FSteps[11].ExpectRuntimeHeld := TRUE;
FSteps[11].CheckFinalization := TRUE;
FSteps[11].ExpectedFinalizationCount := 2;
FSteps[11].ExpectedCompletionCount := 2;
FSteps[11].ExpectedFinalResult := E_Result.Passed;
FSteps[11].ExpectedHookCount := 1;
FSteps[11].ExpectedHooks[1].Hook := E_LifecycleHook.Aggregate;
FSteps[11].ExpectedHooks[1].State := E_State.Completed;
FSteps[11].ExpectedHooks[1].Enabled := TRUE;
{endregion}
END_METHOD

END_FUNCTION_BLOCK

// ---- SelfTests/TestCases/TestSuite_TestCaseLifecycle/Test_LifecycleResetError.TcPOU
{region 'Documentation'}
(*!
<summary>Checks Error before CompleteReset finalizes without executing Abort cleanup.</summary>
*)
{endregion}
FUNCTION_BLOCK Test_LifecycleResetError EXTENDS TestCaseLifecycleTestBase

SUPER^();

{region 'Documentation'}
(*!
<summary>Defines explicit exceptional-path stimuli and contract-derived observations.</summary>
*)
{endregion}
METHOD PROTECTED ConfigureScenario
FSubjectPreparationCount := 0;
FSubjectTestCount := 1;
FStepCount := 2;

{region "01 - Reset fails before completion"}
// Report Error inside ProcessReset before acknowledging completion.
// Expect Completing with Error; subsequent ProcessAbort must be called disabled, not as cleanup.
FSteps[1].RequestReset := TRUE;
FSteps[1].ResetError := TRUE;
FSteps[1].ExpectedState := E_State.Completing;
FSteps[1].ExpectedResult := E_Result.Error;
FSteps[1].ExpectedReady := FALSE;
FSteps[1].ExpectedPassedCount := 0;
FSteps[1].ExpectedFailedCount := 0;
FSteps[1].ExpectedHookCount := 6;
FSteps[1].ExpectedHooks[1].Hook := E_LifecycleHook.Reset;
FSteps[1].ExpectedHooks[1].State := E_State.Reset;
FSteps[1].ExpectedHooks[1].Enabled := TRUE;
FSteps[1].ExpectedHooks[2].Hook := E_LifecycleHook.Abort;
FSteps[1].ExpectedHooks[2].State := E_State.Completing;
FSteps[1].ExpectedHooks[2].Enabled := FALSE;
FSteps[1].ExpectedHooks[3].Hook := E_LifecycleHook.Preparations;
FSteps[1].ExpectedHooks[3].State := E_State.Completing;
FSteps[1].ExpectedHooks[3].Enabled := FALSE;
FSteps[1].ExpectedHooks[4].Hook := E_LifecycleHook.Tests;
FSteps[1].ExpectedHooks[4].State := E_State.Completing;
FSteps[1].ExpectedHooks[4].Enabled := FALSE;
FSteps[1].ExpectedHooks[5].Hook := E_LifecycleHook.Assertions;
FSteps[1].ExpectedHooks[5].State := E_State.Completing;
FSteps[1].ExpectedHooks[5].Enabled := FALSE;
FSteps[1].ExpectedHooks[6].Hook := E_LifecycleHook.Aggregate;
FSteps[1].ExpectedHooks[6].State := E_State.Completing;
FSteps[1].ExpectedHooks[6].Enabled := TRUE;
{endregion}

{region "02 - Observe terminal Error without Abort"}
// The following call reaches Completed; only aggregation remains in the recorded processing
// hooks.
FSteps[2].ExpectedState := E_State.Completed;
FSteps[2].ExpectedResult := E_Result.Error;
FSteps[2].ExpectedReady := FALSE;
FSteps[2].ExpectedPassedCount := 0;
FSteps[2].ExpectedFailedCount := 0;
FSteps[2].ExpectedHookCount := 1;
FSteps[2].ExpectedHooks[1].Hook := E_LifecycleHook.Aggregate;
FSteps[2].ExpectedHooks[1].State := E_State.Completed;
FSteps[2].ExpectedHooks[1].Enabled := TRUE;
{endregion}
END_METHOD

END_FUNCTION_BLOCK

// ---- SelfTests/TestCases/TestSuite_TestCaseLifecycle/Test_LifecycleResetTimeout.TcPOU
{region 'Documentation'}
(*!
<summary>Withholds CompleteReset and verifies direct timeout finalization without Abort processing.</summary>
*)
{endregion}
FUNCTION_BLOCK Test_LifecycleResetTimeout EXTENDS TestCaseLifecycleTestBase

SUPER^();

{region 'Documentation'}
(*!
<summary>Defines explicit exceptional-path stimuli and contract-derived observations.</summary>
*)
{endregion}
METHOD PROTECTED ConfigureScenario
// Exercise the real cyclic timer; these checkpoints check the timeout path and retained flag,
// not an exact elapsed-time boundary. The outer Test Case timeout bounds a missing transition.
FSubjectPreparationCount := 0;
FSubjectTestCount := 1;
FStepCount := 9;
FSubjectConfig.ResetTimeout := T#50ms;

{region "01 - Request Reset and hold acknowledgement"}
// Request Reset once and withhold its completion acknowledgement.
FSteps[1].RequestReset := TRUE;
FSteps[1].ResetCompleted := FALSE;
FSteps[1].ExpectedState := E_State.Reset;
FSteps[1].ExpectedResult := E_Result.NotEvaluated;
FSteps[1].ExpectedReady := FALSE;
FSteps[1].ExpectedPassedCount := 0;
FSteps[1].ExpectedFailedCount := 0;
FSteps[1].ExpectedHookCount := 6;
FSteps[1].ExpectedHooks[1].Hook := E_LifecycleHook.Reset;
FSteps[1].ExpectedHooks[1].State := E_State.Reset;
FSteps[1].ExpectedHooks[1].Enabled := TRUE;
FSteps[1].ExpectedHooks[2].Hook := E_LifecycleHook.Abort;
FSteps[1].ExpectedHooks[2].State := E_State.Reset;
FSteps[1].ExpectedHooks[2].Enabled := FALSE;
FSteps[1].ExpectedHooks[3].Hook := E_LifecycleHook.Preparations;
FSteps[1].ExpectedHooks[3].State := E_State.Reset;
FSteps[1].ExpectedHooks[3].Enabled := FALSE;
FSteps[1].ExpectedHooks[4].Hook := E_LifecycleHook.Tests;
FSteps[1].ExpectedHooks[4].State := E_State.Reset;
FSteps[1].ExpectedHooks[4].Enabled := FALSE;
FSteps[1].ExpectedHooks[5].Hook := E_LifecycleHook.Assertions;
FSteps[1].ExpectedHooks[5].State := E_State.Reset;
FSteps[1].ExpectedHooks[5].Enabled := FALSE;
FSteps[1].ExpectedHooks[6].Hook := E_LifecycleHook.Aggregate;
FSteps[1].ExpectedHooks[6].State := E_State.Reset;
FSteps[1].ExpectedHooks[6].Enabled := TRUE;
{endregion}

{region "02 - Wait for Reset timeout without Abort"}
// Keep reset acknowledgement withheld while repeating this checkpoint.
// Timeout must reach Completing with Error directly, without active Abort cleanup.
FSteps[2].WaitForTransition := TRUE;
FSteps[2].WaitingState := E_State.Reset;
FSteps[2].ResetCompleted := FALSE;
FSteps[2].ExpectedResetTimeout := TRUE;
FSteps[2].ExpectedState := E_State.Completing;
FSteps[2].ExpectedResult := E_Result.Error;
FSteps[2].ExpectedReady := FALSE;
FSteps[2].ExpectedPassedCount := 0;
FSteps[2].ExpectedFailedCount := 0;
FSteps[2].ExpectedHookCount := 5;
FSteps[2].ExpectedHooks[1].Hook := E_LifecycleHook.Abort;
FSteps[2].ExpectedHooks[1].State := E_State.Completing;
FSteps[2].ExpectedHooks[1].Enabled := FALSE;
FSteps[2].ExpectedHooks[2].Hook := E_LifecycleHook.Preparations;
FSteps[2].ExpectedHooks[2].State := E_State.Completing;
FSteps[2].ExpectedHooks[2].Enabled := FALSE;
FSteps[2].ExpectedHooks[3].Hook := E_LifecycleHook.Tests;
FSteps[2].ExpectedHooks[3].State := E_State.Completing;
FSteps[2].ExpectedHooks[3].Enabled := FALSE;
FSteps[2].ExpectedHooks[4].Hook := E_LifecycleHook.Assertions;
FSteps[2].ExpectedHooks[4].State := E_State.Completing;
FSteps[2].ExpectedHooks[4].Enabled := FALSE;
FSteps[2].ExpectedHooks[5].Hook := E_LifecycleHook.Aggregate;
FSteps[2].ExpectedHooks[5].State := E_State.Completing;
FSteps[2].ExpectedHooks[5].Enabled := TRUE;
{endregion}

{region "03 - Retain timeout at completion"}
// Reach Completed and retain the Reset-timeout diagnostic.
FSteps[3].ExpectedResetTimeout := TRUE;
FSteps[3].ExpectedState := E_State.Completed;
FSteps[3].ExpectedResult := E_Result.Error;
FSteps[3].ExpectedReady := FALSE;
FSteps[3].ExpectedPassedCount := 0;
FSteps[3].ExpectedFailedCount := 0;
FSteps[3].ExpectedHookCount := 1;
FSteps[3].ExpectedHooks[1].Hook := E_LifecycleHook.Aggregate;
FSteps[3].ExpectedHooks[1].State := E_State.Completed;
FSteps[3].ExpectedHooks[1].Enabled := TRUE;
{endregion}

{region "04 - Reset clears held timeout and result"}
FSteps[4].ExpectedState := E_State.Idle;
FSteps[4].ExpectedResult := E_Result.NotEvaluated;
FSteps[4].ExpectedReady := TRUE;
FSteps[4].ExpectedPassedCount := 0;
FSteps[4].ExpectedFailedCount := 0;
FSteps[4].CheckFinalization := TRUE;
FSteps[4].ExpectedFinalizationCount := 1;
FSteps[4].ExpectedCompletionCount := 1;
FSteps[4].ExpectedFinalResult := E_Result.Error;
FSteps[4].RequestReset := TRUE;
FSteps[4].PreparationTargetReached := TRUE;
FSteps[4].ExpectRuntimeCleared := TRUE;
FSteps[4].ExpectedHookCount := 6;
FSteps[4].ExpectedHooks[1].Hook := E_LifecycleHook.Reset;
FSteps[4].ExpectedHooks[1].State := E_State.Reset;
FSteps[4].ExpectedHooks[1].Enabled := TRUE;
FSteps[4].ExpectedHooks[2].Hook := E_LifecycleHook.Abort;
FSteps[4].ExpectedHooks[2].State := E_State.Idle;
FSteps[4].ExpectedHooks[2].Enabled := FALSE;
FSteps[4].ExpectedHooks[3].Hook := E_LifecycleHook.Preparations;
FSteps[4].ExpectedHooks[3].State := E_State.Idle;
FSteps[4].ExpectedHooks[3].Enabled := FALSE;
FSteps[4].ExpectedHooks[4].Hook := E_LifecycleHook.Tests;
FSteps[4].ExpectedHooks[4].State := E_State.Idle;
FSteps[4].ExpectedHooks[4].Enabled := FALSE;
FSteps[4].ExpectedHooks[5].Hook := E_LifecycleHook.Assertions;
FSteps[4].ExpectedHooks[5].State := E_State.Idle;
FSteps[4].ExpectedHooks[5].Enabled := FALSE;
FSteps[4].ExpectedHooks[6].Hook := E_LifecycleHook.Aggregate;
FSteps[4].ExpectedHooks[6].State := E_State.Idle;
FSteps[4].ExpectedHooks[6].Enabled := TRUE;
{endregion}

{region "05 - Start after timeout recovery"}
FSteps[5].ExpectedState := E_State.Starting;
FSteps[5].ExpectedResult := E_Result.NotEvaluated;
FSteps[5].ExpectedReady := FALSE;
FSteps[5].ExpectedPassedCount := 0;
FSteps[5].ExpectedFailedCount := 0;
FSteps[5].CheckFinalization := TRUE;
FSteps[5].ExpectedFinalizationCount := 1;
FSteps[5].ExpectedCompletionCount := 1;
FSteps[5].ExpectedFinalResult := E_Result.Error;
FSteps[5].RequestStart := TRUE;
FSteps[5].PreparationTargetReached := TRUE;
FSteps[5].ExpectedHookCount := 5;
FSteps[5].ExpectedHooks[1].Hook := E_LifecycleHook.Abort;
FSteps[5].ExpectedHooks[1].State := E_State.Starting;
FSteps[5].ExpectedHooks[1].Enabled := FALSE;
FSteps[5].ExpectedHooks[2].Hook := E_LifecycleHook.Preparations;
FSteps[5].ExpectedHooks[2].State := E_State.Starting;
FSteps[5].ExpectedHooks[2].Enabled := FALSE;
FSteps[5].ExpectedHooks[3].Hook := E_LifecycleHook.Tests;
FSteps[5].ExpectedHooks[3].State := E_State.Starting;
FSteps[5].ExpectedHooks[3].Enabled := FALSE;
FSteps[5].ExpectedHooks[4].Hook := E_LifecycleHook.Assertions;
FSteps[5].ExpectedHooks[4].State := E_State.Starting;
FSteps[5].ExpectedHooks[4].Enabled := FALSE;
FSteps[5].ExpectedHooks[5].Hook := E_LifecycleHook.Aggregate;
FSteps[5].ExpectedHooks[5].State := E_State.Starting;
FSteps[5].ExpectedHooks[5].Enabled := TRUE;
{endregion}

{region "06 - Execute without previous timeout flags"}
FSteps[6].ExpectedState := E_State.Running;
FSteps[6].ExpectedResult := E_Result.NotEvaluated;
FSteps[6].ExpectedReady := FALSE;
FSteps[6].ExpectedPassedCount := 2;
FSteps[6].ExpectedFailedCount := 0;
FSteps[6].CheckFinalization := TRUE;
FSteps[6].ExpectedFinalizationCount := 1;
FSteps[6].ExpectedCompletionCount := 1;
FSteps[6].ExpectedFinalResult := E_Result.Error;
FSteps[6].ExpectedHookCount := 5;
FSteps[6].ExpectedHooks[1].Hook := E_LifecycleHook.Abort;
FSteps[6].ExpectedHooks[1].State := E_State.Running;
FSteps[6].ExpectedHooks[1].Enabled := FALSE;
FSteps[6].ExpectedHooks[2].Hook := E_LifecycleHook.Preparations;
FSteps[6].ExpectedHooks[2].State := E_State.Running;
FSteps[6].ExpectedHooks[2].Enabled := FALSE;
FSteps[6].ExpectedHooks[3].Hook := E_LifecycleHook.Tests;
FSteps[6].ExpectedHooks[3].State := E_State.Running;
FSteps[6].ExpectedHooks[3].Enabled := TRUE;
FSteps[6].ExpectedHooks[4].Hook := E_LifecycleHook.Assertions;
FSteps[6].ExpectedHooks[4].State := E_State.Running;
FSteps[6].ExpectedHooks[4].Enabled := TRUE;
FSteps[6].ExpectedHooks[5].Hook := E_LifecycleHook.Aggregate;
FSteps[6].ExpectedHooks[5].State := E_State.Running;
FSteps[6].ExpectedHooks[5].Enabled := TRUE;
{endregion}

{region "07 - Finalize the recovered run"}
FSteps[7].ExpectedState := E_State.Completing;
FSteps[7].ExpectedResult := E_Result.Passed;
FSteps[7].ExpectedReady := FALSE;
FSteps[7].ExpectedPassedCount := 2;
FSteps[7].ExpectedFailedCount := 0;
FSteps[7].FinishTests := TRUE;
FSteps[7].CheckFinalization := TRUE;
FSteps[7].ExpectedFinalizationCount := 2;
FSteps[7].ExpectedCompletionCount := 1;
FSteps[7].ExpectedFinalResult := E_Result.Passed;
FSteps[7].ExpectedHookCount := 5;
FSteps[7].ExpectedHooks[1].Hook := E_LifecycleHook.Abort;
FSteps[7].ExpectedHooks[1].State := E_State.Running;
FSteps[7].ExpectedHooks[1].Enabled := FALSE;
FSteps[7].ExpectedHooks[2].Hook := E_LifecycleHook.Preparations;
FSteps[7].ExpectedHooks[2].State := E_State.Running;
FSteps[7].ExpectedHooks[2].Enabled := FALSE;
FSteps[7].ExpectedHooks[3].Hook := E_LifecycleHook.Tests;
FSteps[7].ExpectedHooks[3].State := E_State.Running;
FSteps[7].ExpectedHooks[3].Enabled := TRUE;
FSteps[7].ExpectedHooks[4].Hook := E_LifecycleHook.Assertions;
FSteps[7].ExpectedHooks[4].State := E_State.Completing;
FSteps[7].ExpectedHooks[4].Enabled := FALSE;
FSteps[7].ExpectedHooks[5].Hook := E_LifecycleHook.Aggregate;
FSteps[7].ExpectedHooks[5].State := E_State.Completing;
FSteps[7].ExpectedHooks[5].Enabled := TRUE;
{endregion}

{region "08 - Complete the recovered run"}
FSteps[8].ExpectedState := E_State.Completed;
FSteps[8].ExpectedResult := E_Result.Passed;
FSteps[8].ExpectedReady := FALSE;
FSteps[8].ExpectedPassedCount := 2;
FSteps[8].ExpectedFailedCount := 0;
FSteps[8].ExpectRuntimeHeld := TRUE;
FSteps[8].CheckFinalization := TRUE;
FSteps[8].ExpectedFinalizationCount := 2;
FSteps[8].ExpectedCompletionCount := 2;
FSteps[8].ExpectedFinalResult := E_Result.Passed;
FSteps[8].ExpectedHookCount := 1;
FSteps[8].ExpectedHooks[1].Hook := E_LifecycleHook.Aggregate;
FSteps[8].ExpectedHooks[1].State := E_State.Completed;
FSteps[8].ExpectedHooks[1].Enabled := TRUE;
{endregion}

{region "09 - Hold the recovered completion without new events"}
FSteps[9].ExpectedState := E_State.Completed;
FSteps[9].ExpectedResult := E_Result.Passed;
FSteps[9].ExpectedReady := FALSE;
FSteps[9].ExpectedPassedCount := 2;
FSteps[9].ExpectedFailedCount := 0;
FSteps[9].ExpectQuietCall := TRUE;
FSteps[9].ExpectRuntimeHeld := TRUE;
FSteps[9].CheckFinalization := TRUE;
FSteps[9].ExpectedFinalizationCount := 2;
FSteps[9].ExpectedCompletionCount := 2;
FSteps[9].ExpectedFinalResult := E_Result.Passed;
FSteps[9].ExpectedHookCount := 1;
FSteps[9].ExpectedHooks[1].Hook := E_LifecycleHook.Aggregate;
FSteps[9].ExpectedHooks[1].State := E_State.Completed;
FSteps[9].ExpectedHooks[1].Enabled := TRUE;
{endregion}
END_METHOD

END_FUNCTION_BLOCK

// ---- SelfTests/TestCases/TestSuite_TestCaseLifecycle/Test_LifecycleResetDuringExecution.TcPOU
{region 'Documentation'}
(*!
<summary>Checks Reset interruption of an active run, including request priority and cleared child results.</summary>
*)
{endregion}
FUNCTION_BLOCK Test_LifecycleResetDuringExecution EXTENDS TestCaseLifecycleTestBase

SUPER^();

{region 'Documentation'}
(*!
<summary>Defines explicit exceptional-path stimuli and contract-derived observations.</summary>
*)
{endregion}
METHOD PROTECTED ConfigureScenario
FSubjectPreparationCount := 0;
FSubjectTestCount := 1;
FStepCount := 9;

{region "01 - Reset to Idle"}
// Establish Idle through the parent Reset request; both child results must be cleared.
FSteps[1].RequestReset := TRUE;
FSteps[1].ExpectedState := E_State.Idle;
FSteps[1].ExpectedResult := E_Result.NotEvaluated;
FSteps[1].ExpectedReady := TRUE;
FSteps[1].ExpectedPassedCount := 0;
FSteps[1].ExpectedFailedCount := 0;
FSteps[1].ExpectedHookCount := 6;
FSteps[1].ExpectedHooks[1].Hook := E_LifecycleHook.Reset;
FSteps[1].ExpectedHooks[1].State := E_State.Reset;
FSteps[1].ExpectedHooks[1].Enabled := TRUE;
FSteps[1].ExpectedHooks[2].Hook := E_LifecycleHook.Abort;
FSteps[1].ExpectedHooks[2].State := E_State.Idle;
FSteps[1].ExpectedHooks[2].Enabled := FALSE;
FSteps[1].ExpectedHooks[3].Hook := E_LifecycleHook.Preparations;
FSteps[1].ExpectedHooks[3].State := E_State.Idle;
FSteps[1].ExpectedHooks[3].Enabled := FALSE;
FSteps[1].ExpectedHooks[4].Hook := E_LifecycleHook.Tests;
FSteps[1].ExpectedHooks[4].State := E_State.Idle;
FSteps[1].ExpectedHooks[4].Enabled := FALSE;
FSteps[1].ExpectedHooks[5].Hook := E_LifecycleHook.Assertions;
FSteps[1].ExpectedHooks[5].State := E_State.Idle;
FSteps[1].ExpectedHooks[5].Enabled := FALSE;
FSteps[1].ExpectedHooks[6].Hook := E_LifecycleHook.Aggregate;
FSteps[1].ExpectedHooks[6].State := E_State.Idle;
FSteps[1].ExpectedHooks[6].Enabled := TRUE;
{endregion}

{region "02 - Accept Start"}
// Accept Start into Starting; processing and Assertion evaluation are not active yet.
FSteps[2].RequestStart := TRUE;
FSteps[2].ExpectedState := E_State.Starting;
FSteps[2].ExpectedResult := E_Result.NotEvaluated;
FSteps[2].ExpectedReady := FALSE;
FSteps[2].ExpectedPassedCount := 0;
FSteps[2].ExpectedFailedCount := 0;
FSteps[2].ExpectedHookCount := 5;
FSteps[2].ExpectedHooks[1].Hook := E_LifecycleHook.Abort;
FSteps[2].ExpectedHooks[1].State := E_State.Starting;
FSteps[2].ExpectedHooks[1].Enabled := FALSE;
FSteps[2].ExpectedHooks[2].Hook := E_LifecycleHook.Preparations;
FSteps[2].ExpectedHooks[2].State := E_State.Starting;
FSteps[2].ExpectedHooks[2].Enabled := FALSE;
FSteps[2].ExpectedHooks[3].Hook := E_LifecycleHook.Tests;
FSteps[2].ExpectedHooks[3].State := E_State.Starting;
FSteps[2].ExpectedHooks[3].Enabled := FALSE;
FSteps[2].ExpectedHooks[4].Hook := E_LifecycleHook.Assertions;
FSteps[2].ExpectedHooks[4].State := E_State.Starting;
FSteps[2].ExpectedHooks[4].Enabled := FALSE;
FSteps[2].ExpectedHooks[5].Hook := E_LifecycleHook.Aggregate;
FSteps[2].ExpectedHooks[5].State := E_State.Starting;
FSteps[2].ExpectedHooks[5].Enabled := TRUE;
{endregion}

{region "03 - Establish active execution"}
// Enter Running and evaluate both children; owner Result stays NotEvaluated until finalization.
FSteps[3].ExpectedState := E_State.Running;
FSteps[3].ExpectedResult := E_Result.NotEvaluated;
FSteps[3].ExpectedReady := FALSE;
FSteps[3].ExpectedPassedCount := 2;
FSteps[3].ExpectedFailedCount := 0;
FSteps[3].ExpectedHookCount := 5;
FSteps[3].ExpectedHooks[1].Hook := E_LifecycleHook.Abort;
FSteps[3].ExpectedHooks[1].State := E_State.Running;
FSteps[3].ExpectedHooks[1].Enabled := FALSE;
FSteps[3].ExpectedHooks[2].Hook := E_LifecycleHook.Preparations;
FSteps[3].ExpectedHooks[2].State := E_State.Running;
FSteps[3].ExpectedHooks[2].Enabled := FALSE;
FSteps[3].ExpectedHooks[3].Hook := E_LifecycleHook.Tests;
FSteps[3].ExpectedHooks[3].State := E_State.Running;
FSteps[3].ExpectedHooks[3].Enabled := TRUE;
FSteps[3].ExpectedHooks[4].Hook := E_LifecycleHook.Assertions;
FSteps[3].ExpectedHooks[4].State := E_State.Running;
FSteps[3].ExpectedHooks[4].Enabled := TRUE;
FSteps[3].ExpectedHooks[5].Hook := E_LifecycleHook.Aggregate;
FSteps[3].ExpectedHooks[5].State := E_State.Running;
FSteps[3].ExpectedHooks[5].Enabled := TRUE;
{endregion}

{region "04 - Reset wins competing requests"}
// Submit Reset, Abort and Start together during Running.
// Reset must win, clear child results and finish in Idle without active Abort cleanup.
FSteps[4].RequestReset := TRUE;
FSteps[4].RequestAbort := TRUE;
FSteps[4].RequestStart := TRUE;
FSteps[4].ExpectedState := E_State.Idle;
FSteps[4].ExpectedResult := E_Result.NotEvaluated;
FSteps[4].ExpectedReady := TRUE;
FSteps[4].ExpectedPassedCount := 0;
FSteps[4].ExpectedFailedCount := 0;
FSteps[4].ExpectedHookCount := 6;
FSteps[4].ExpectedHooks[1].Hook := E_LifecycleHook.Reset;
FSteps[4].ExpectedHooks[1].State := E_State.Reset;
FSteps[4].ExpectedHooks[1].Enabled := TRUE;
FSteps[4].ExpectedHooks[2].Hook := E_LifecycleHook.Abort;
FSteps[4].ExpectedHooks[2].State := E_State.Idle;
FSteps[4].ExpectedHooks[2].Enabled := FALSE;
FSteps[4].ExpectedHooks[3].Hook := E_LifecycleHook.Preparations;
FSteps[4].ExpectedHooks[3].State := E_State.Idle;
FSteps[4].ExpectedHooks[3].Enabled := FALSE;
FSteps[4].ExpectedHooks[4].Hook := E_LifecycleHook.Tests;
FSteps[4].ExpectedHooks[4].State := E_State.Idle;
FSteps[4].ExpectedHooks[4].Enabled := FALSE;
FSteps[4].ExpectedHooks[5].Hook := E_LifecycleHook.Assertions;
FSteps[4].ExpectedHooks[5].State := E_State.Idle;
FSteps[4].ExpectedHooks[5].Enabled := FALSE;
FSteps[4].ExpectedHooks[6].Hook := E_LifecycleHook.Aggregate;
FSteps[4].ExpectedHooks[6].State := E_State.Idle;
FSteps[4].ExpectedHooks[6].Enabled := TRUE;
{endregion}

{region "05 - No deferred automatic Start"}
// Stay Idle after the competing requests were consumed; Start must not survive the Reset.
FSteps[5].ExpectedState := E_State.Idle;
FSteps[5].ExpectedResult := E_Result.NotEvaluated;
FSteps[5].ExpectedReady := TRUE;
FSteps[5].ExpectedPassedCount := 0;
FSteps[5].ExpectedFailedCount := 0;
FSteps[5].ExpectedHookCount := 5;
FSteps[5].ExpectedHooks[1].Hook := E_LifecycleHook.Abort;
FSteps[5].ExpectedHooks[1].State := E_State.Idle;
FSteps[5].ExpectedHooks[1].Enabled := FALSE;
FSteps[5].ExpectedHooks[2].Hook := E_LifecycleHook.Preparations;
FSteps[5].ExpectedHooks[2].State := E_State.Idle;
FSteps[5].ExpectedHooks[2].Enabled := FALSE;
FSteps[5].ExpectedHooks[3].Hook := E_LifecycleHook.Tests;
FSteps[5].ExpectedHooks[3].State := E_State.Idle;
FSteps[5].ExpectedHooks[3].Enabled := FALSE;
FSteps[5].ExpectedHooks[4].Hook := E_LifecycleHook.Assertions;
FSteps[5].ExpectedHooks[4].State := E_State.Idle;
FSteps[5].ExpectedHooks[4].Enabled := FALSE;
FSteps[5].ExpectedHooks[5].Hook := E_LifecycleHook.Aggregate;
FSteps[5].ExpectedHooks[5].State := E_State.Idle;
FSteps[5].ExpectedHooks[5].Enabled := TRUE;
{endregion}

{region "06 - Accept fresh Start"}
// Only this fresh Start may begin another execution.
FSteps[6].RequestStart := TRUE;
FSteps[6].ExpectedState := E_State.Starting;
FSteps[6].ExpectedResult := E_Result.NotEvaluated;
FSteps[6].ExpectedReady := FALSE;
FSteps[6].ExpectedPassedCount := 0;
FSteps[6].ExpectedFailedCount := 0;
FSteps[6].ExpectedHookCount := 5;
FSteps[6].ExpectedHooks[1].Hook := E_LifecycleHook.Abort;
FSteps[6].ExpectedHooks[1].State := E_State.Starting;
FSteps[6].ExpectedHooks[1].Enabled := FALSE;
FSteps[6].ExpectedHooks[2].Hook := E_LifecycleHook.Preparations;
FSteps[6].ExpectedHooks[2].State := E_State.Starting;
FSteps[6].ExpectedHooks[2].Enabled := FALSE;
FSteps[6].ExpectedHooks[3].Hook := E_LifecycleHook.Tests;
FSteps[6].ExpectedHooks[3].State := E_State.Starting;
FSteps[6].ExpectedHooks[3].Enabled := FALSE;
FSteps[6].ExpectedHooks[4].Hook := E_LifecycleHook.Assertions;
FSteps[6].ExpectedHooks[4].State := E_State.Starting;
FSteps[6].ExpectedHooks[4].Enabled := FALSE;
FSteps[6].ExpectedHooks[5].Hook := E_LifecycleHook.Aggregate;
FSteps[6].ExpectedHooks[5].State := E_State.Starting;
FSteps[6].ExpectedHooks[5].Enabled := TRUE;
{endregion}

{region "07 - Execute after Reset"}
// Enter Running and evaluate both children; owner Result stays NotEvaluated until finalization.
FSteps[7].ExpectedState := E_State.Running;
FSteps[7].ExpectedResult := E_Result.NotEvaluated;
FSteps[7].ExpectedReady := FALSE;
FSteps[7].ExpectedPassedCount := 2;
FSteps[7].ExpectedFailedCount := 0;
FSteps[7].ExpectedHookCount := 5;
FSteps[7].ExpectedHooks[1].Hook := E_LifecycleHook.Abort;
FSteps[7].ExpectedHooks[1].State := E_State.Running;
FSteps[7].ExpectedHooks[1].Enabled := FALSE;
FSteps[7].ExpectedHooks[2].Hook := E_LifecycleHook.Preparations;
FSteps[7].ExpectedHooks[2].State := E_State.Running;
FSteps[7].ExpectedHooks[2].Enabled := FALSE;
FSteps[7].ExpectedHooks[3].Hook := E_LifecycleHook.Tests;
FSteps[7].ExpectedHooks[3].State := E_State.Running;
FSteps[7].ExpectedHooks[3].Enabled := TRUE;
FSteps[7].ExpectedHooks[4].Hook := E_LifecycleHook.Assertions;
FSteps[7].ExpectedHooks[4].State := E_State.Running;
FSteps[7].ExpectedHooks[4].Enabled := TRUE;
FSteps[7].ExpectedHooks[5].Hook := E_LifecycleHook.Aggregate;
FSteps[7].ExpectedHooks[5].State := E_State.Running;
FSteps[7].ExpectedHooks[5].Enabled := TRUE;
{endregion}

{region "08 - Complete inside test processing"}
// CompleteTests changes phase inside ProcessTests; subsequent Assertions must already be
// disabled.
FSteps[8].FinishTests := TRUE;
FSteps[8].ExpectedState := E_State.Completing;
FSteps[8].ExpectedResult := E_Result.Passed;
FSteps[8].ExpectedReady := FALSE;
FSteps[8].ExpectedPassedCount := 2;
FSteps[8].ExpectedFailedCount := 0;
FSteps[8].ExpectedHookCount := 5;
FSteps[8].ExpectedHooks[1].Hook := E_LifecycleHook.Abort;
FSteps[8].ExpectedHooks[1].State := E_State.Running;
FSteps[8].ExpectedHooks[1].Enabled := FALSE;
FSteps[8].ExpectedHooks[2].Hook := E_LifecycleHook.Preparations;
FSteps[8].ExpectedHooks[2].State := E_State.Running;
FSteps[8].ExpectedHooks[2].Enabled := FALSE;
FSteps[8].ExpectedHooks[3].Hook := E_LifecycleHook.Tests;
FSteps[8].ExpectedHooks[3].State := E_State.Running;
FSteps[8].ExpectedHooks[3].Enabled := TRUE;
FSteps[8].ExpectedHooks[4].Hook := E_LifecycleHook.Assertions;
FSteps[8].ExpectedHooks[4].State := E_State.Completing;
FSteps[8].ExpectedHooks[4].Enabled := FALSE;
FSteps[8].ExpectedHooks[5].Hook := E_LifecycleHook.Aggregate;
FSteps[8].ExpectedHooks[5].State := E_State.Completing;
FSteps[8].ExpectedHooks[5].Enabled := TRUE;
{endregion}

{region "09 - Observe terminal completion"}
// The following call reaches Completed; only aggregation remains in the recorded processing
// hooks.
FSteps[9].ExpectedState := E_State.Completed;
FSteps[9].ExpectedResult := E_Result.Passed;
FSteps[9].ExpectedReady := FALSE;
FSteps[9].ExpectedPassedCount := 2;
FSteps[9].ExpectedFailedCount := 0;
FSteps[9].ExpectedHookCount := 1;
FSteps[9].ExpectedHooks[1].Hook := E_LifecycleHook.Aggregate;
FSteps[9].ExpectedHooks[1].State := E_State.Completed;
FSteps[9].ExpectedHooks[1].Enabled := TRUE;
{endregion}
END_METHOD

END_FUNCTION_BLOCK

// ---- SelfTests/TestCases/TestSuite_TestCaseLifecycle/Test_LifecycleFailedToError.TcPOU
{region 'Documentation'}
(*!
<summary>Checks that a Failed child cannot suppress a later owner Error and controlled cleanup.</summary>
*)
{endregion}
FUNCTION_BLOCK Test_LifecycleFailedToError EXTENDS TestCaseLifecycleTestBase

SUPER^();

{region 'Documentation'}
(*!
<summary>Defines explicit exceptional-path stimuli and contract-derived observations.</summary>
*)
{endregion}
METHOD PROTECTED ConfigureScenario
FSubjectPreparationCount := 0;
FSubjectTestCount := 1;
FStepCount := 6;

{region "01 - Reset to Idle"}
// Establish Idle through the parent Reset request; both child results must be cleared.
FSteps[1].RequestReset := TRUE;
FSteps[1].ExpectedState := E_State.Idle;
FSteps[1].ExpectedResult := E_Result.NotEvaluated;
FSteps[1].ExpectedReady := TRUE;
FSteps[1].ExpectedPassedCount := 0;
FSteps[1].ExpectedFailedCount := 0;
FSteps[1].ExpectedHookCount := 6;
FSteps[1].ExpectedHooks[1].Hook := E_LifecycleHook.Reset;
FSteps[1].ExpectedHooks[1].State := E_State.Reset;
FSteps[1].ExpectedHooks[1].Enabled := TRUE;
FSteps[1].ExpectedHooks[2].Hook := E_LifecycleHook.Abort;
FSteps[1].ExpectedHooks[2].State := E_State.Idle;
FSteps[1].ExpectedHooks[2].Enabled := FALSE;
FSteps[1].ExpectedHooks[3].Hook := E_LifecycleHook.Preparations;
FSteps[1].ExpectedHooks[3].State := E_State.Idle;
FSteps[1].ExpectedHooks[3].Enabled := FALSE;
FSteps[1].ExpectedHooks[4].Hook := E_LifecycleHook.Tests;
FSteps[1].ExpectedHooks[4].State := E_State.Idle;
FSteps[1].ExpectedHooks[4].Enabled := FALSE;
FSteps[1].ExpectedHooks[5].Hook := E_LifecycleHook.Assertions;
FSteps[1].ExpectedHooks[5].State := E_State.Idle;
FSteps[1].ExpectedHooks[5].Enabled := FALSE;
FSteps[1].ExpectedHooks[6].Hook := E_LifecycleHook.Aggregate;
FSteps[1].ExpectedHooks[6].State := E_State.Idle;
FSteps[1].ExpectedHooks[6].Enabled := TRUE;
{endregion}

{region "02 - Accept Start"}
// Accept Start into Starting; processing and Assertion evaluation are not active yet.
FSteps[2].RequestStart := TRUE;
FSteps[2].ExpectedState := E_State.Starting;
FSteps[2].ExpectedResult := E_Result.NotEvaluated;
FSteps[2].ExpectedReady := FALSE;
FSteps[2].ExpectedPassedCount := 0;
FSteps[2].ExpectedFailedCount := 0;
FSteps[2].ExpectedHookCount := 5;
FSteps[2].ExpectedHooks[1].Hook := E_LifecycleHook.Abort;
FSteps[2].ExpectedHooks[1].State := E_State.Starting;
FSteps[2].ExpectedHooks[1].Enabled := FALSE;
FSteps[2].ExpectedHooks[2].Hook := E_LifecycleHook.Preparations;
FSteps[2].ExpectedHooks[2].State := E_State.Starting;
FSteps[2].ExpectedHooks[2].Enabled := FALSE;
FSteps[2].ExpectedHooks[3].Hook := E_LifecycleHook.Tests;
FSteps[2].ExpectedHooks[3].State := E_State.Starting;
FSteps[2].ExpectedHooks[3].Enabled := FALSE;
FSteps[2].ExpectedHooks[4].Hook := E_LifecycleHook.Assertions;
FSteps[2].ExpectedHooks[4].State := E_State.Starting;
FSteps[2].ExpectedHooks[4].Enabled := FALSE;
FSteps[2].ExpectedHooks[5].Hook := E_LifecycleHook.Aggregate;
FSteps[2].ExpectedHooks[5].State := E_State.Starting;
FSteps[2].ExpectedHooks[5].Enabled := TRUE;
{endregion}

{region "03 - Establish a child failure"}
// First produce a real child failure; the companion Assertion still passes.
FSteps[3].AssertionCondition := FALSE;
FSteps[3].ExpectedState := E_State.Running;
FSteps[3].ExpectedResult := E_Result.NotEvaluated;
FSteps[3].ExpectedReady := FALSE;
FSteps[3].ExpectedPassedCount := 1;
FSteps[3].ExpectedFailedCount := 1;
FSteps[3].ExpectedHookCount := 5;
FSteps[3].ExpectedHooks[1].Hook := E_LifecycleHook.Abort;
FSteps[3].ExpectedHooks[1].State := E_State.Running;
FSteps[3].ExpectedHooks[1].Enabled := FALSE;
FSteps[3].ExpectedHooks[2].Hook := E_LifecycleHook.Preparations;
FSteps[3].ExpectedHooks[2].State := E_State.Running;
FSteps[3].ExpectedHooks[2].Enabled := FALSE;
FSteps[3].ExpectedHooks[3].Hook := E_LifecycleHook.Tests;
FSteps[3].ExpectedHooks[3].State := E_State.Running;
FSteps[3].ExpectedHooks[3].Enabled := TRUE;
FSteps[3].ExpectedHooks[4].Hook := E_LifecycleHook.Assertions;
FSteps[3].ExpectedHooks[4].State := E_State.Running;
FSteps[3].ExpectedHooks[4].Enabled := TRUE;
FSteps[3].ExpectedHooks[5].Hook := E_LifecycleHook.Aggregate;
FSteps[3].ExpectedHooks[5].State := E_State.Running;
FSteps[3].ExpectedHooks[5].Enabled := TRUE;
{endregion}

{region "04 - Escalate framework error during tests"}
// Raise a framework Error from ProcessTests despite the existing Failed child.
// ProcessAbort ran disabled earlier in this call; cleanup starts on the following call.
FSteps[4].TestError := TRUE;
FSteps[4].ExpectedState := E_State.AbortingFromError;
FSteps[4].ExpectedResult := E_Result.Error;
FSteps[4].ExpectedReady := FALSE;
FSteps[4].ExpectedPassedCount := 1;
FSteps[4].ExpectedFailedCount := 1;
FSteps[4].ExpectedHookCount := 5;
FSteps[4].ExpectedHooks[1].Hook := E_LifecycleHook.Abort;
FSteps[4].ExpectedHooks[1].State := E_State.Running;
FSteps[4].ExpectedHooks[1].Enabled := FALSE;
FSteps[4].ExpectedHooks[2].Hook := E_LifecycleHook.Preparations;
FSteps[4].ExpectedHooks[2].State := E_State.Running;
FSteps[4].ExpectedHooks[2].Enabled := FALSE;
FSteps[4].ExpectedHooks[3].Hook := E_LifecycleHook.Tests;
FSteps[4].ExpectedHooks[3].State := E_State.Running;
FSteps[4].ExpectedHooks[3].Enabled := TRUE;
FSteps[4].ExpectedHooks[4].Hook := E_LifecycleHook.Assertions;
FSteps[4].ExpectedHooks[4].State := E_State.AbortingFromError;
FSteps[4].ExpectedHooks[4].Enabled := FALSE;
FSteps[4].ExpectedHooks[5].Hook := E_LifecycleHook.Aggregate;
FSteps[4].ExpectedHooks[5].State := E_State.AbortingFromError;
FSteps[4].ExpectedHooks[5].Enabled := TRUE;
{endregion}

{region "05 - Complete error-abort cleanup"}
// Now execute error-abort cleanup and acknowledge it; finalization must retain Error.
FSteps[5].ExpectedState := E_State.Completing;
FSteps[5].ExpectedResult := E_Result.Error;
FSteps[5].ExpectedReady := FALSE;
FSteps[5].ExpectedPassedCount := 1;
FSteps[5].ExpectedFailedCount := 1;
FSteps[5].ExpectedHookCount := 5;
FSteps[5].ExpectedHooks[1].Hook := E_LifecycleHook.Abort;
FSteps[5].ExpectedHooks[1].State := E_State.AbortingFromError;
FSteps[5].ExpectedHooks[1].Enabled := TRUE;
FSteps[5].ExpectedHooks[2].Hook := E_LifecycleHook.Preparations;
FSteps[5].ExpectedHooks[2].State := E_State.Completing;
FSteps[5].ExpectedHooks[2].Enabled := FALSE;
FSteps[5].ExpectedHooks[3].Hook := E_LifecycleHook.Tests;
FSteps[5].ExpectedHooks[3].State := E_State.Completing;
FSteps[5].ExpectedHooks[3].Enabled := FALSE;
FSteps[5].ExpectedHooks[4].Hook := E_LifecycleHook.Assertions;
FSteps[5].ExpectedHooks[4].State := E_State.Completing;
FSteps[5].ExpectedHooks[4].Enabled := FALSE;
FSteps[5].ExpectedHooks[5].Hook := E_LifecycleHook.Aggregate;
FSteps[5].ExpectedHooks[5].State := E_State.Completing;
FSteps[5].ExpectedHooks[5].Enabled := TRUE;
{endregion}

{region "06 - Observe terminal Error"}
// The following call reaches Completed; only aggregation remains in the recorded processing
// hooks.
FSteps[6].ExpectedState := E_State.Completed;
FSteps[6].ExpectedResult := E_Result.Error;
FSteps[6].ExpectedReady := FALSE;
FSteps[6].ExpectedPassedCount := 1;
FSteps[6].ExpectedFailedCount := 1;
FSteps[6].ExpectedHookCount := 1;
FSteps[6].ExpectedHooks[1].Hook := E_LifecycleHook.Aggregate;
FSteps[6].ExpectedHooks[1].State := E_State.Completed;
FSteps[6].ExpectedHooks[1].Enabled := TRUE;
{endregion}
END_METHOD

END_FUNCTION_BLOCK

// ---- SelfTests/TestCases/TestSuite_TestCaseLifecycle/Test_LifecycleInvalidTestAdvance.TcPOU
{region 'Documentation'}
(*!
<summary>Checks an out-of-range NextTestState call escalates without entering an unconfigured state.</summary>
*)
{endregion}
FUNCTION_BLOCK Test_LifecycleInvalidTestAdvance EXTENDS TestCaseLifecycleTestBase

SUPER^();

{region 'Documentation'}
(*!
<summary>Defines explicit exceptional-path stimuli and contract-derived observations.</summary>
*)
{endregion}
METHOD PROTECTED ConfigureScenario
FSubjectPreparationCount := 0;
FSubjectTestCount := 1;
FStepCount := 6;

{region "01 - Reset to Idle"}
// Establish Idle through the parent Reset request; both child results must be cleared.
FSteps[1].RequestReset := TRUE;
FSteps[1].ExpectedState := E_State.Idle;
FSteps[1].ExpectedResult := E_Result.NotEvaluated;
FSteps[1].ExpectedReady := TRUE;
FSteps[1].ExpectedPassedCount := 0;
FSteps[1].ExpectedFailedCount := 0;
FSteps[1].ExpectedHookCount := 6;
FSteps[1].ExpectedHooks[1].Hook := E_LifecycleHook.Reset;
FSteps[1].ExpectedHooks[1].State := E_State.Reset;
FSteps[1].ExpectedHooks[1].Enabled := TRUE;
FSteps[1].ExpectedHooks[2].Hook := E_LifecycleHook.Abort;
FSteps[1].ExpectedHooks[2].State := E_State.Idle;
FSteps[1].ExpectedHooks[2].Enabled := FALSE;
FSteps[1].ExpectedHooks[3].Hook := E_LifecycleHook.Preparations;
FSteps[1].ExpectedHooks[3].State := E_State.Idle;
FSteps[1].ExpectedHooks[3].Enabled := FALSE;
FSteps[1].ExpectedHooks[4].Hook := E_LifecycleHook.Tests;
FSteps[1].ExpectedHooks[4].State := E_State.Idle;
FSteps[1].ExpectedHooks[4].Enabled := FALSE;
FSteps[1].ExpectedHooks[5].Hook := E_LifecycleHook.Assertions;
FSteps[1].ExpectedHooks[5].State := E_State.Idle;
FSteps[1].ExpectedHooks[5].Enabled := FALSE;
FSteps[1].ExpectedHooks[6].Hook := E_LifecycleHook.Aggregate;
FSteps[1].ExpectedHooks[6].State := E_State.Idle;
FSteps[1].ExpectedHooks[6].Enabled := TRUE;
{endregion}

{region "02 - Accept Start"}
// Accept Start into Starting; processing and Assertion evaluation are not active yet.
FSteps[2].RequestStart := TRUE;
FSteps[2].ExpectedState := E_State.Starting;
FSteps[2].ExpectedResult := E_Result.NotEvaluated;
FSteps[2].ExpectedReady := FALSE;
FSteps[2].ExpectedPassedCount := 0;
FSteps[2].ExpectedFailedCount := 0;
FSteps[2].ExpectedHookCount := 5;
FSteps[2].ExpectedHooks[1].Hook := E_LifecycleHook.Abort;
FSteps[2].ExpectedHooks[1].State := E_State.Starting;
FSteps[2].ExpectedHooks[1].Enabled := FALSE;
FSteps[2].ExpectedHooks[2].Hook := E_LifecycleHook.Preparations;
FSteps[2].ExpectedHooks[2].State := E_State.Starting;
FSteps[2].ExpectedHooks[2].Enabled := FALSE;
FSteps[2].ExpectedHooks[3].Hook := E_LifecycleHook.Tests;
FSteps[2].ExpectedHooks[3].State := E_State.Starting;
FSteps[2].ExpectedHooks[3].Enabled := FALSE;
FSteps[2].ExpectedHooks[4].Hook := E_LifecycleHook.Assertions;
FSteps[2].ExpectedHooks[4].State := E_State.Starting;
FSteps[2].ExpectedHooks[4].Enabled := FALSE;
FSteps[2].ExpectedHooks[5].Hook := E_LifecycleHook.Aggregate;
FSteps[2].ExpectedHooks[5].State := E_State.Starting;
FSteps[2].ExpectedHooks[5].Enabled := TRUE;
{endregion}

{region "03 - Enter only configured Test state"}
// Enter Running and evaluate both children; owner Result stays NotEvaluated until finalization.
FSteps[3].ExpectedState := E_State.Running;
FSteps[3].ExpectedResult := E_Result.NotEvaluated;
FSteps[3].ExpectedReady := FALSE;
FSteps[3].ExpectedPassedCount := 2;
FSteps[3].ExpectedFailedCount := 0;
FSteps[3].ExpectedHookCount := 5;
FSteps[3].ExpectedHooks[1].Hook := E_LifecycleHook.Abort;
FSteps[3].ExpectedHooks[1].State := E_State.Running;
FSteps[3].ExpectedHooks[1].Enabled := FALSE;
FSteps[3].ExpectedHooks[2].Hook := E_LifecycleHook.Preparations;
FSteps[3].ExpectedHooks[2].State := E_State.Running;
FSteps[3].ExpectedHooks[2].Enabled := FALSE;
FSteps[3].ExpectedHooks[3].Hook := E_LifecycleHook.Tests;
FSteps[3].ExpectedHooks[3].State := E_State.Running;
FSteps[3].ExpectedHooks[3].Enabled := TRUE;
FSteps[3].ExpectedHooks[4].Hook := E_LifecycleHook.Assertions;
FSteps[3].ExpectedHooks[4].State := E_State.Running;
FSteps[3].ExpectedHooks[4].Enabled := TRUE;
FSteps[3].ExpectedHooks[5].Hook := E_LifecycleHook.Aggregate;
FSteps[3].ExpectedHooks[5].State := E_State.Running;
FSteps[3].ExpectedHooks[5].Enabled := TRUE;
{endregion}

{region "04 - Reject Test-state overrun"}
// Advance beyond the only configured Test state.
// Reject the request with Error; later hooks see AbortingFromError and Assertions are disabled.
FSteps[4].AdvanceTest := TRUE;
FSteps[4].ExpectedState := E_State.AbortingFromError;
FSteps[4].ExpectedResult := E_Result.Error;
FSteps[4].ExpectedReady := FALSE;
FSteps[4].ExpectedPassedCount := 2;
FSteps[4].ExpectedFailedCount := 0;
FSteps[4].ExpectedHookCount := 5;
FSteps[4].ExpectedHooks[1].Hook := E_LifecycleHook.Abort;
FSteps[4].ExpectedHooks[1].State := E_State.Running;
FSteps[4].ExpectedHooks[1].Enabled := FALSE;
FSteps[4].ExpectedHooks[2].Hook := E_LifecycleHook.Preparations;
FSteps[4].ExpectedHooks[2].State := E_State.Running;
FSteps[4].ExpectedHooks[2].Enabled := FALSE;
FSteps[4].ExpectedHooks[3].Hook := E_LifecycleHook.Tests;
FSteps[4].ExpectedHooks[3].State := E_State.Running;
FSteps[4].ExpectedHooks[3].Enabled := TRUE;
FSteps[4].ExpectedHooks[4].Hook := E_LifecycleHook.Assertions;
FSteps[4].ExpectedHooks[4].State := E_State.AbortingFromError;
FSteps[4].ExpectedHooks[4].Enabled := FALSE;
FSteps[4].ExpectedHooks[5].Hook := E_LifecycleHook.Aggregate;
FSteps[4].ExpectedHooks[5].State := E_State.AbortingFromError;
FSteps[4].ExpectedHooks[5].Enabled := TRUE;
{endregion}

{region "05 - Complete error-abort cleanup"}
// Execute the pending error-abort cleanup on the following call, then finalize with Error.
FSteps[5].ExpectedState := E_State.Completing;
FSteps[5].ExpectedResult := E_Result.Error;
FSteps[5].ExpectedReady := FALSE;
FSteps[5].ExpectedPassedCount := 2;
FSteps[5].ExpectedFailedCount := 0;
FSteps[5].ExpectedHookCount := 5;
FSteps[5].ExpectedHooks[1].Hook := E_LifecycleHook.Abort;
FSteps[5].ExpectedHooks[1].State := E_State.AbortingFromError;
FSteps[5].ExpectedHooks[1].Enabled := TRUE;
FSteps[5].ExpectedHooks[2].Hook := E_LifecycleHook.Preparations;
FSteps[5].ExpectedHooks[2].State := E_State.Completing;
FSteps[5].ExpectedHooks[2].Enabled := FALSE;
FSteps[5].ExpectedHooks[3].Hook := E_LifecycleHook.Tests;
FSteps[5].ExpectedHooks[3].State := E_State.Completing;
FSteps[5].ExpectedHooks[3].Enabled := FALSE;
FSteps[5].ExpectedHooks[4].Hook := E_LifecycleHook.Assertions;
FSteps[5].ExpectedHooks[4].State := E_State.Completing;
FSteps[5].ExpectedHooks[4].Enabled := FALSE;
FSteps[5].ExpectedHooks[5].Hook := E_LifecycleHook.Aggregate;
FSteps[5].ExpectedHooks[5].State := E_State.Completing;
FSteps[5].ExpectedHooks[5].Enabled := TRUE;
{endregion}

{region "06 - Observe terminal Error"}
// The following call reaches Completed; only aggregation remains in the recorded processing
// hooks.
FSteps[6].ExpectedState := E_State.Completed;
FSteps[6].ExpectedResult := E_Result.Error;
FSteps[6].ExpectedReady := FALSE;
FSteps[6].ExpectedPassedCount := 2;
FSteps[6].ExpectedFailedCount := 0;
FSteps[6].ExpectedHookCount := 1;
FSteps[6].ExpectedHooks[1].Hook := E_LifecycleHook.Aggregate;
FSteps[6].ExpectedHooks[1].State := E_State.Completed;
FSteps[6].ExpectedHooks[1].Enabled := TRUE;
{endregion}
END_METHOD

END_FUNCTION_BLOCK

// ---- SelfTests/TestCases/TestSuite_TestCaseLifecycle/Test_LifecycleInvalidPreparationTransition.TcPOU
{region 'Documentation'}
(*!
<summary>Rejects completion before the Preparation target is reached; no Test hook may become enabled.</summary>
*)
{endregion}
FUNCTION_BLOCK Test_LifecycleInvalidPreparationTransition EXTENDS TestCaseLifecycleTestBase

SUPER^();

{region 'Documentation'}
(*!
<summary>Defines explicit exceptional-path stimuli and contract-derived observations.</summary>
*)
{endregion}
METHOD PROTECTED ConfigureScenario
FSubjectPreparationCount := 1;
FSubjectTestCount := 1;
FStepCount := 6;

{region "01 - Reset to Idle"}
// Establish Idle through the parent Reset request; both child results must be cleared.
FSteps[1].RequestReset := TRUE;
FSteps[1].ExpectedState := E_State.Idle;
FSteps[1].ExpectedResult := E_Result.NotEvaluated;
FSteps[1].ExpectedReady := TRUE;
FSteps[1].ExpectedPassedCount := 0;
FSteps[1].ExpectedFailedCount := 0;
FSteps[1].ExpectedHookCount := 6;
FSteps[1].ExpectedHooks[1].Hook := E_LifecycleHook.Reset;
FSteps[1].ExpectedHooks[1].State := E_State.Reset;
FSteps[1].ExpectedHooks[1].Enabled := TRUE;
FSteps[1].ExpectedHooks[2].Hook := E_LifecycleHook.Abort;
FSteps[1].ExpectedHooks[2].State := E_State.Idle;
FSteps[1].ExpectedHooks[2].Enabled := FALSE;
FSteps[1].ExpectedHooks[3].Hook := E_LifecycleHook.Preparations;
FSteps[1].ExpectedHooks[3].State := E_State.Idle;
FSteps[1].ExpectedHooks[3].Enabled := FALSE;
FSteps[1].ExpectedHooks[4].Hook := E_LifecycleHook.Tests;
FSteps[1].ExpectedHooks[4].State := E_State.Idle;
FSteps[1].ExpectedHooks[4].Enabled := FALSE;
FSteps[1].ExpectedHooks[5].Hook := E_LifecycleHook.Assertions;
FSteps[1].ExpectedHooks[5].State := E_State.Idle;
FSteps[1].ExpectedHooks[5].Enabled := FALSE;
FSteps[1].ExpectedHooks[6].Hook := E_LifecycleHook.Aggregate;
FSteps[1].ExpectedHooks[6].State := E_State.Idle;
FSteps[1].ExpectedHooks[6].Enabled := TRUE;
{endregion}

{region "02 - Accept Start"}
// Accept Start into Starting; processing and Assertion evaluation are not active yet.
FSteps[2].RequestStart := TRUE;
FSteps[2].ExpectedState := E_State.Starting;
FSteps[2].ExpectedResult := E_Result.NotEvaluated;
FSteps[2].ExpectedReady := FALSE;
FSteps[2].ExpectedPassedCount := 0;
FSteps[2].ExpectedFailedCount := 0;
FSteps[2].ExpectedHookCount := 5;
FSteps[2].ExpectedHooks[1].Hook := E_LifecycleHook.Abort;
FSteps[2].ExpectedHooks[1].State := E_State.Starting;
FSteps[2].ExpectedHooks[1].Enabled := FALSE;
FSteps[2].ExpectedHooks[2].Hook := E_LifecycleHook.Preparations;
FSteps[2].ExpectedHooks[2].State := E_State.Starting;
FSteps[2].ExpectedHooks[2].Enabled := FALSE;
FSteps[2].ExpectedHooks[3].Hook := E_LifecycleHook.Tests;
FSteps[2].ExpectedHooks[3].State := E_State.Starting;
FSteps[2].ExpectedHooks[3].Enabled := FALSE;
FSteps[2].ExpectedHooks[4].Hook := E_LifecycleHook.Assertions;
FSteps[2].ExpectedHooks[4].State := E_State.Starting;
FSteps[2].ExpectedHooks[4].Enabled := FALSE;
FSteps[2].ExpectedHooks[5].Hook := E_LifecycleHook.Aggregate;
FSteps[2].ExpectedHooks[5].State := E_State.Starting;
FSteps[2].ExpectedHooks[5].Enabled := TRUE;
{endregion}

{region "03 - Wait for target"}
// Enter Preparing without evaluating Assertions; the target has not been reached.
FSteps[3].ExpectedState := E_State.Preparing;
FSteps[3].ExpectedResult := E_Result.NotEvaluated;
FSteps[3].ExpectedReady := FALSE;
FSteps[3].ExpectedPassedCount := 0;
FSteps[3].ExpectedFailedCount := 0;
FSteps[3].ExpectedHookCount := 5;
FSteps[3].ExpectedHooks[1].Hook := E_LifecycleHook.Abort;
FSteps[3].ExpectedHooks[1].State := E_State.Preparing;
FSteps[3].ExpectedHooks[1].Enabled := FALSE;
FSteps[3].ExpectedHooks[2].Hook := E_LifecycleHook.Preparations;
FSteps[3].ExpectedHooks[2].State := E_State.Preparing;
FSteps[3].ExpectedHooks[2].Enabled := TRUE;
FSteps[3].ExpectedHooks[3].Hook := E_LifecycleHook.Tests;
FSteps[3].ExpectedHooks[3].State := E_State.Preparing;
FSteps[3].ExpectedHooks[3].Enabled := FALSE;
FSteps[3].ExpectedHooks[4].Hook := E_LifecycleHook.Assertions;
FSteps[3].ExpectedHooks[4].State := E_State.Preparing;
FSteps[3].ExpectedHooks[4].Enabled := FALSE;
FSteps[3].ExpectedHooks[5].Hook := E_LifecycleHook.Aggregate;
FSteps[3].ExpectedHooks[5].State := E_State.Preparing;
FSteps[3].ExpectedHooks[5].Enabled := TRUE;
{endregion}

{region "04 - Reject premature completion"}
// Call CompletePreparations without a reached target.
// Reject the transition, latch Error and remain Preparing for the rest of this call.
FSteps[4].FinishPreparations := TRUE;
FSteps[4].ExpectedState := E_State.Preparing;
FSteps[4].ExpectedResult := E_Result.Error;
FSteps[4].ExpectedReady := FALSE;
FSteps[4].ExpectedPassedCount := 0;
FSteps[4].ExpectedFailedCount := 0;
FSteps[4].ExpectedHookCount := 5;
FSteps[4].ExpectedHooks[1].Hook := E_LifecycleHook.Abort;
FSteps[4].ExpectedHooks[1].State := E_State.Preparing;
FSteps[4].ExpectedHooks[1].Enabled := FALSE;
FSteps[4].ExpectedHooks[2].Hook := E_LifecycleHook.Preparations;
FSteps[4].ExpectedHooks[2].State := E_State.Preparing;
FSteps[4].ExpectedHooks[2].Enabled := TRUE;
FSteps[4].ExpectedHooks[3].Hook := E_LifecycleHook.Tests;
FSteps[4].ExpectedHooks[3].State := E_State.Preparing;
FSteps[4].ExpectedHooks[3].Enabled := FALSE;
FSteps[4].ExpectedHooks[4].Hook := E_LifecycleHook.Assertions;
FSteps[4].ExpectedHooks[4].State := E_State.Preparing;
FSteps[4].ExpectedHooks[4].Enabled := FALSE;
FSteps[4].ExpectedHooks[5].Hook := E_LifecycleHook.Aggregate;
FSteps[4].ExpectedHooks[5].State := E_State.Preparing;
FSteps[4].ExpectedHooks[5].Enabled := TRUE;
{endregion}

{region "05 - Finalize through error cleanup"}
// The following Sequencer routes the held Error through active abort cleanup to Completing.
FSteps[5].ExpectedState := E_State.Completing;
FSteps[5].ExpectedResult := E_Result.Error;
FSteps[5].ExpectedReady := FALSE;
FSteps[5].ExpectedPassedCount := 0;
FSteps[5].ExpectedFailedCount := 0;
FSteps[5].ExpectedHookCount := 5;
FSteps[5].ExpectedHooks[1].Hook := E_LifecycleHook.Abort;
FSteps[5].ExpectedHooks[1].State := E_State.AbortingFromError;
FSteps[5].ExpectedHooks[1].Enabled := TRUE;
FSteps[5].ExpectedHooks[2].Hook := E_LifecycleHook.Preparations;
FSteps[5].ExpectedHooks[2].State := E_State.Completing;
FSteps[5].ExpectedHooks[2].Enabled := FALSE;
FSteps[5].ExpectedHooks[3].Hook := E_LifecycleHook.Tests;
FSteps[5].ExpectedHooks[3].State := E_State.Completing;
FSteps[5].ExpectedHooks[3].Enabled := FALSE;
FSteps[5].ExpectedHooks[4].Hook := E_LifecycleHook.Assertions;
FSteps[5].ExpectedHooks[4].State := E_State.Completing;
FSteps[5].ExpectedHooks[4].Enabled := FALSE;
FSteps[5].ExpectedHooks[5].Hook := E_LifecycleHook.Aggregate;
FSteps[5].ExpectedHooks[5].State := E_State.Completing;
FSteps[5].ExpectedHooks[5].Enabled := TRUE;
{endregion}

{region "06 - Observe terminal Error"}
// The following call reaches Completed; only aggregation remains in the recorded processing
// hooks.
FSteps[6].ExpectedState := E_State.Completed;
FSteps[6].ExpectedResult := E_Result.Error;
FSteps[6].ExpectedReady := FALSE;
FSteps[6].ExpectedPassedCount := 0;
FSteps[6].ExpectedFailedCount := 0;
FSteps[6].ExpectedHookCount := 1;
FSteps[6].ExpectedHooks[1].Hook := E_LifecycleHook.Aggregate;
FSteps[6].ExpectedHooks[1].State := E_State.Completed;
FSteps[6].ExpectedHooks[1].Enabled := TRUE;
{endregion}
END_METHOD

END_FUNCTION_BLOCK

// ---- SelfTests/TestCases/TestSuite_TestCaseLifecycle/Test_LifecycleRepeatAfterPassed.TcPOU
{region 'Documentation'}
(*!
<summary>Checks stable Passed completion, one-shot finalization and a fresh successful run after Reset.</summary>
*)
{endregion}
FUNCTION_BLOCK Test_LifecycleRepeatAfterPassed EXTENDS TestCaseLifecycleTestBase

SUPER^();

{region 'Documentation'}
(*!
<summary>Defines two independent run outcomes and cumulative event expectations across Reset.</summary>
*)
{endregion}
METHOD PROTECTED ConfigureScenario
FSubjectPreparationCount := 0;
FSubjectTestCount := 1;
FStepCount := 15;

{region "01 - Reset establishes the initial Idle state"}
FSteps[1].ExpectedState := E_State.Idle;
FSteps[1].ExpectedResult := E_Result.NotEvaluated;
FSteps[1].ExpectedReady := TRUE;
FSteps[1].ExpectedPassedCount := 0;
FSteps[1].ExpectedFailedCount := 0;
FSteps[1].RequestReset := TRUE;
FSteps[1].ExpectRuntimeCleared := TRUE;
FSteps[1].CheckFinalization := TRUE;
FSteps[1].ExpectedFinalizationCount := 0;
FSteps[1].ExpectedCompletionCount := 0;
FSteps[1].ExpectedFinalResult := E_Result.Passed;
FSteps[1].ExpectedHookCount := 6;
FSteps[1].ExpectedHooks[1].Hook := E_LifecycleHook.Reset;
FSteps[1].ExpectedHooks[1].State := E_State.Reset;
FSteps[1].ExpectedHooks[1].Enabled := TRUE;
FSteps[1].ExpectedHooks[2].Hook := E_LifecycleHook.Abort;
FSteps[1].ExpectedHooks[2].State := E_State.Idle;
FSteps[1].ExpectedHooks[2].Enabled := FALSE;
FSteps[1].ExpectedHooks[3].Hook := E_LifecycleHook.Preparations;
FSteps[1].ExpectedHooks[3].State := E_State.Idle;
FSteps[1].ExpectedHooks[3].Enabled := FALSE;
FSteps[1].ExpectedHooks[4].Hook := E_LifecycleHook.Tests;
FSteps[1].ExpectedHooks[4].State := E_State.Idle;
FSteps[1].ExpectedHooks[4].Enabled := FALSE;
FSteps[1].ExpectedHooks[5].Hook := E_LifecycleHook.Assertions;
FSteps[1].ExpectedHooks[5].State := E_State.Idle;
FSteps[1].ExpectedHooks[5].Enabled := FALSE;
FSteps[1].ExpectedHooks[6].Hook := E_LifecycleHook.Aggregate;
FSteps[1].ExpectedHooks[6].State := E_State.Idle;
FSteps[1].ExpectedHooks[6].Enabled := TRUE;
{endregion}

{region "02 - Start the first execution"}
FSteps[2].ExpectedState := E_State.Starting;
FSteps[2].ExpectedResult := E_Result.NotEvaluated;
FSteps[2].ExpectedReady := FALSE;
FSteps[2].ExpectedPassedCount := 0;
FSteps[2].ExpectedFailedCount := 0;
FSteps[2].RequestStart := TRUE;
FSteps[2].CheckFinalization := TRUE;
FSteps[2].ExpectedFinalizationCount := 0;
FSteps[2].ExpectedCompletionCount := 0;
FSteps[2].ExpectedFinalResult := E_Result.Passed;
FSteps[2].ExpectedHookCount := 5;
FSteps[2].ExpectedHooks[1].Hook := E_LifecycleHook.Abort;
FSteps[2].ExpectedHooks[1].State := E_State.Starting;
FSteps[2].ExpectedHooks[1].Enabled := FALSE;
FSteps[2].ExpectedHooks[2].Hook := E_LifecycleHook.Preparations;
FSteps[2].ExpectedHooks[2].State := E_State.Starting;
FSteps[2].ExpectedHooks[2].Enabled := FALSE;
FSteps[2].ExpectedHooks[3].Hook := E_LifecycleHook.Tests;
FSteps[2].ExpectedHooks[3].State := E_State.Starting;
FSteps[2].ExpectedHooks[3].Enabled := FALSE;
FSteps[2].ExpectedHooks[4].Hook := E_LifecycleHook.Assertions;
FSteps[2].ExpectedHooks[4].State := E_State.Starting;
FSteps[2].ExpectedHooks[4].Enabled := FALSE;
FSteps[2].ExpectedHooks[5].Hook := E_LifecycleHook.Aggregate;
FSteps[2].ExpectedHooks[5].State := E_State.Starting;
FSteps[2].ExpectedHooks[5].Enabled := TRUE;
{endregion}

{region "03 - Evaluate both child Assertions"}
FSteps[3].ExpectedState := E_State.Running;
FSteps[3].ExpectedResult := E_Result.NotEvaluated;
FSteps[3].ExpectedReady := FALSE;
FSteps[3].ExpectedPassedCount := 2;
FSteps[3].ExpectedFailedCount := 0;
FSteps[3].AssertionCondition := TRUE;
FSteps[3].CheckFinalization := TRUE;
FSteps[3].ExpectedFinalizationCount := 0;
FSteps[3].ExpectedCompletionCount := 0;
FSteps[3].ExpectedFinalResult := E_Result.Passed;
FSteps[3].ExpectedHookCount := 5;
FSteps[3].ExpectedHooks[1].Hook := E_LifecycleHook.Abort;
FSteps[3].ExpectedHooks[1].State := E_State.Running;
FSteps[3].ExpectedHooks[1].Enabled := FALSE;
FSteps[3].ExpectedHooks[2].Hook := E_LifecycleHook.Preparations;
FSteps[3].ExpectedHooks[2].State := E_State.Running;
FSteps[3].ExpectedHooks[2].Enabled := FALSE;
FSteps[3].ExpectedHooks[3].Hook := E_LifecycleHook.Tests;
FSteps[3].ExpectedHooks[3].State := E_State.Running;
FSteps[3].ExpectedHooks[3].Enabled := TRUE;
FSteps[3].ExpectedHooks[4].Hook := E_LifecycleHook.Assertions;
FSteps[3].ExpectedHooks[4].State := E_State.Running;
FSteps[3].ExpectedHooks[4].Enabled := TRUE;
FSteps[3].ExpectedHooks[5].Hook := E_LifecycleHook.Aggregate;
FSteps[3].ExpectedHooks[5].State := E_State.Running;
FSteps[3].ExpectedHooks[5].Enabled := TRUE;
{endregion}

{region "04 - Finalize the first result"}
FSteps[4].ExpectedState := E_State.Completing;
FSteps[4].ExpectedResult := E_Result.Passed;
FSteps[4].ExpectedReady := FALSE;
FSteps[4].ExpectedPassedCount := 2;
FSteps[4].ExpectedFailedCount := 0;
FSteps[4].FinishTests := TRUE;
FSteps[4].CheckFinalization := TRUE;
FSteps[4].ExpectedFinalizationCount := 1;
FSteps[4].ExpectedCompletionCount := 0;
FSteps[4].ExpectedFinalResult := E_Result.Passed;
FSteps[4].ExpectedHookCount := 5;
FSteps[4].ExpectedHooks[1].Hook := E_LifecycleHook.Abort;
FSteps[4].ExpectedHooks[1].State := E_State.Running;
FSteps[4].ExpectedHooks[1].Enabled := FALSE;
FSteps[4].ExpectedHooks[2].Hook := E_LifecycleHook.Preparations;
FSteps[4].ExpectedHooks[2].State := E_State.Running;
FSteps[4].ExpectedHooks[2].Enabled := FALSE;
FSteps[4].ExpectedHooks[3].Hook := E_LifecycleHook.Tests;
FSteps[4].ExpectedHooks[3].State := E_State.Running;
FSteps[4].ExpectedHooks[3].Enabled := TRUE;
FSteps[4].ExpectedHooks[4].Hook := E_LifecycleHook.Assertions;
FSteps[4].ExpectedHooks[4].State := E_State.Completing;
FSteps[4].ExpectedHooks[4].Enabled := FALSE;
FSteps[4].ExpectedHooks[5].Hook := E_LifecycleHook.Aggregate;
FSteps[4].ExpectedHooks[5].State := E_State.Completing;
FSteps[4].ExpectedHooks[5].Enabled := TRUE;
{endregion}

{region "05 - Observe the final Completed transition"}
FSteps[5].ExpectedState := E_State.Completed;
FSteps[5].ExpectedResult := E_Result.Passed;
FSteps[5].ExpectedReady := FALSE;
FSteps[5].ExpectedPassedCount := 2;
FSteps[5].ExpectedFailedCount := 0;
FSteps[5].CheckFinalization := TRUE;
FSteps[5].ExpectedFinalizationCount := 1;
FSteps[5].ExpectedCompletionCount := 1;
FSteps[5].ExpectedFinalResult := E_Result.Passed;
FSteps[5].ExpectRuntimeHeld := TRUE;
FSteps[5].ExpectedHookCount := 1;
FSteps[5].ExpectedHooks[1].Hook := E_LifecycleHook.Aggregate;
FSteps[5].ExpectedHooks[1].State := E_State.Completed;
FSteps[5].ExpectedHooks[1].Enabled := TRUE;
{endregion}

{region "06 - Ignore processing inputs while Completed"}
FSteps[6].ExpectedState := E_State.Completed;
FSteps[6].ExpectedResult := E_Result.Passed;
FSteps[6].ExpectedReady := FALSE;
FSteps[6].ExpectedPassedCount := 2;
FSteps[6].ExpectedFailedCount := 0;
FSteps[6].CheckFinalization := TRUE;
FSteps[6].ExpectedFinalizationCount := 1;
FSteps[6].ExpectedCompletionCount := 1;
FSteps[6].ExpectedFinalResult := E_Result.Passed;
FSteps[6].ExpectRuntimeHeld := TRUE;
FSteps[6].ExpectQuietCall := TRUE;
FSteps[6].Ready := FALSE;
FSteps[6].ResetError := TRUE;
FSteps[6].AbortError := TRUE;
FSteps[6].TestError := TRUE;
FSteps[6].PreparationError := TRUE;
FSteps[6].AdvancePreparation := TRUE;
FSteps[6].FinishPreparations := TRUE;
FSteps[6].AdvanceTest := TRUE;
FSteps[6].FinishTests := TRUE;
FSteps[6].AssertionCondition := FALSE;
FSteps[6].ExpectedHookCount := 1;
FSteps[6].ExpectedHooks[1].Hook := E_LifecycleHook.Aggregate;
FSteps[6].ExpectedHooks[1].State := E_State.Completed;
FSteps[6].ExpectedHooks[1].Enabled := TRUE;
{endregion}

